	E_CELL_MANAGER_STATE.WAIT_GRIPPER1_CONTENT:
		IF rtOperatorChoice.Q AND xOperatorChoiceAllowed THEN
			IF uiOperatorChoice = UINT#1 THEN
				IF Config.uiTypeCount = UINT#1 THEN
					uiBlankPayloadType := UINT#1;
					IF xPrestartGripper2Occupied THEN
						eState := E_CELL_MANAGER_STATE.WAIT_GRIPPER2_CONTENT;
					ELSE
						xSafetyHomeRequired := FALSE;
						xStoppedPoseValid := FALSE;
						xRunning := TRUE;
						eState := E_CELL_MANAGER_STATE.PLAN_TARGET;
					END_IF;
				ELSE
					eState := E_CELL_MANAGER_STATE.WAIT_GRIPPER1_TYPE;
				END_IF;
			ELSIF uiOperatorChoice = UINT#2 THEN
				Diag.stWarning.uiCode := WRN_GRIPPER1_CONTENT;
				Diag.stWarning.udiSequence := Diag.stWarning.udiSequence + UDINT#1;
				IF Diag.stWarning.udiSequence = UDINT#0 THEN Diag.stWarning.udiSequence := UDINT#1; END_IF;
				eState := E_CELL_MANAGER_STATE.IDLE;
			ELSE
				Diag.stWarning.uiCode := WRN_OPERATOR_REPLY_REJECTED;
				Diag.stWarning.udiSequence := Diag.stWarning.udiSequence + UDINT#1;
				IF Diag.stWarning.udiSequence = UDINT#0 THEN Diag.stWarning.udiSequence := UDINT#1; END_IF;
				eState := E_CELL_MANAGER_STATE.IDLE;
			END_IF;
		END_IF;

	E_CELL_MANAGER_STATE.WAIT_GRIPPER1_TYPE:
		IF rtOperatorChoice.Q AND xOperatorChoiceAllowed THEN
			IF (uiOperatorChoice >= UINT#1)
			AND (uiOperatorChoice <= Config.uiTypeCount) THEN
				uiBlankPayloadType := uiOperatorChoice;
				IF xPrestartGripper2Occupied THEN
					eState := E_CELL_MANAGER_STATE.WAIT_GRIPPER2_CONTENT;
				ELSE
					xSafetyHomeRequired := FALSE;
					xStoppedPoseValid := FALSE;
					xRunning := TRUE;
					eState := E_CELL_MANAGER_STATE.PLAN_TARGET;
				END_IF;
			ELSE
				Diag.stWarning.uiCode := WRN_PAYLOAD_TYPE_CHOICE;
				Diag.stWarning.udiSequence := Diag.stWarning.udiSequence + UDINT#1;
				IF Diag.stWarning.udiSequence = UDINT#0 THEN Diag.stWarning.udiSequence := UDINT#1; END_IF;
				eState := E_CELL_MANAGER_STATE.IDLE;
			END_IF;
		END_IF;

	E_CELL_MANAGER_STATE.WAIT_GRIPPER2_CONTENT:
		IF rtOperatorChoice.Q AND xOperatorChoiceAllowed THEN
			IF uiOperatorChoice = UINT#2 THEN
				IF Config.uiTypeCount = UINT#1 THEN
					uiDetailPayloadType := UINT#1;
				ELSE
					eState := E_CELL_MANAGER_STATE.WAIT_GRIPPER2_TYPE;
				END_IF;
				IF (Config.uiTypeCount = UINT#1) AND xPrestartGripper1Occupied THEN
					IF uiOperatorMachineMask <> UINT#0 THEN
						eState := E_CELL_MANAGER_STATE.WAIT_START_MACHINE;
					ELSE
						// Нет пустого совместимого станка: это не тупик. После
						// идентификации обоих грузов планировщик сначала уложит деталь.
						xSafetyHomeRequired := FALSE;
						xStoppedPoseValid := FALSE;
						xRunning := TRUE;
						eState := E_CELL_MANAGER_STATE.PLAN_TARGET;
					END_IF;
				ELSIF Config.uiTypeCount = UINT#1 THEN
					xSafetyHomeRequired := FALSE;
					xStoppedPoseValid := FALSE;
					xRunning := TRUE;
					eState := E_CELL_MANAGER_STATE.PLAN_TARGET;
				END_IF;
			ELSIF uiOperatorChoice = UINT#1 THEN
				Diag.stWarning.uiCode := WRN_GRIPPER2_CONTENT;
				Diag.stWarning.udiSequence := Diag.stWarning.udiSequence + UDINT#1;
				IF Diag.stWarning.udiSequence = UDINT#0 THEN Diag.stWarning.udiSequence := UDINT#1; END_IF;
				eState := E_CELL_MANAGER_STATE.IDLE;
			ELSE
				Diag.stWarning.uiCode := WRN_OPERATOR_REPLY_REJECTED;
				Diag.stWarning.udiSequence := Diag.stWarning.udiSequence + UDINT#1;
				IF Diag.stWarning.udiSequence = UDINT#0 THEN Diag.stWarning.udiSequence := UDINT#1; END_IF;
				eState := E_CELL_MANAGER_STATE.IDLE;
			END_IF;
		END_IF;

	E_CELL_MANAGER_STATE.WAIT_GRIPPER2_TYPE:
		IF rtOperatorChoice.Q AND xOperatorChoiceAllowed THEN
			IF (uiOperatorChoice >= UINT#1)
			AND (uiOperatorChoice <= Config.uiTypeCount) THEN
				uiDetailPayloadType := uiOperatorChoice;
				IF xPrestartGripper1Occupied THEN
					IF uiOperatorMachineMask <> UINT#0 THEN
						eState := E_CELL_MANAGER_STATE.WAIT_START_MACHINE;
					ELSE
						xSafetyHomeRequired := FALSE;
						xStoppedPoseValid := FALSE;
						xRunning := TRUE;
						eState := E_CELL_MANAGER_STATE.PLAN_TARGET;
					END_IF;
				ELSE
					xSafetyHomeRequired := FALSE;
					xStoppedPoseValid := FALSE;
					xRunning := TRUE;
					eState := E_CELL_MANAGER_STATE.PLAN_TARGET;
				END_IF;
			ELSE
				Diag.stWarning.uiCode := WRN_PAYLOAD_TYPE_CHOICE;
				Diag.stWarning.udiSequence := Diag.stWarning.udiSequence + UDINT#1;
				IF Diag.stWarning.udiSequence = UDINT#0 THEN Diag.stWarning.udiSequence := UDINT#1; END_IF;
				eState := E_CELL_MANAGER_STATE.IDLE;
			END_IF;
		END_IF;

	E_CELL_MANAGER_STATE.WAIT_START_MACHINE:
		IF (uiDetailPayloadType < UINT#1)
		OR (uiDetailPayloadType > Config.uiTypeCount) THEN
			Diag.stWarning.uiCode := WRN_PAYLOAD_TYPE_CHOICE;
			Diag.stWarning.udiSequence := Diag.stWarning.udiSequence + UDINT#1;
			IF Diag.stWarning.udiSequence = UDINT#0 THEN Diag.stWarning.udiSequence := UDINT#1; END_IF;
			eState := E_CELL_MANAGER_STATE.IDLE;
		ELSIF stMagazineStatus.stTypeStatus.aiFreeSlot[uiDetailPayloadType] = SINT#0 THEN
			Diag.stWarning.uiCode := WRN_DETAIL_SLOT_REQUIRED;
			Diag.stWarning.udiSequence := Diag.stWarning.udiSequence + UDINT#1;
			IF Diag.stWarning.udiSequence = UDINT#0 THEN Diag.stWarning.udiSequence := UDINT#1; END_IF;
			eState := E_CELL_MANAGER_STATE.IDLE;
		ELSIF uiOperatorMachineMask = UINT#0 THEN
			// Пока оператор отвечал, пустой станок мог стать недоступен. Сохраняем
			// оба груза и передаём решение общему планировщику вместо отмены старта.
			xSafetyHomeRequired := FALSE;
			xStoppedPoseValid := FALSE;
			xRunning := TRUE;
			eState := E_CELL_MANAGER_STATE.PLAN_TARGET;
		ELSIF rtOperatorChoice.Q AND xOperatorChoiceAllowed THEN
			IF ((uiOperatorChoice = UINT#1) AND ((uiOperatorMachineMask AND UINT#1) <> UINT#0))
			OR ((uiOperatorChoice = UINT#2) AND ((uiOperatorMachineMask AND UINT#2) <> UINT#0))
			OR ((uiOperatorChoice = UINT#3) AND ((uiOperatorMachineMask AND UINT#4) <> UINT#0)) THEN
				uiSelectedMachine := uiOperatorChoice;
				uiSelectedType := uiBlankPayloadType;
				eMachineOperation := E_MACHINE_OPERATION.LOAD;
				xSafetyHomeRequired := FALSE;
				xStoppedPoseValid := FALSE;
				xRunning := TRUE;
				eState := E_CELL_MANAGER_STATE.ROUTE_TO_TARGET;
			ELSE
				Diag.stWarning.uiCode := WRN_START_MACHINE_CHOICE;
				Diag.stWarning.udiSequence := Diag.stWarning.udiSequence + UDINT#1;
				IF Diag.stWarning.udiSequence = UDINT#0 THEN Diag.stWarning.udiSequence := UDINT#1; END_IF;
				eState := E_CELL_MANAGER_STATE.IDLE;
			END_IF;
		END_IF;

	E_CELL_MANAGER_STATE.PLAN_TARGET:
		IF xStopRequested
		AND NOT stRobotStatus.xBusy
		AND NOT stMagazineStatus.xBusy THEN
			xRunning := FALSE;
			eState := E_CELL_MANAGER_STATE.IDLE;

		ELSIF PlanGeometry() THEN
			// Метод зафиксировал резерв или безопасное ожидание свободного ГК.
		ELSIF stRobotStatus.xBlankAvailable
		AND stRobotStatus.xDetailAvailable THEN
			// Два груза после аварийного восстановления — штатная ситуация. Сначала
			// ищем пустой готовый станок строго по типу заготовки. Если загрузить её
			// прямо сейчас некуда, освобождаем захват 2 операцией PUT.
			IF (uiBlankPayloadType < UINT#1)
			OR (uiBlankPayloadType > Config.uiTypeCount) THEN
				Error.dwErrorActive := Error.dwErrorActive OR ERR_MAGAZINE;
				eState := E_CELL_MANAGER_STATE.ERROR;
			ELSIF (uiDetailPayloadType < UINT#1)
			OR (uiDetailPayloadType > Config.uiTypeCount) THEN
				Error.dwErrorActive := Error.dwErrorActive OR ERR_MACHINE;
				eState := E_CELL_MANAGER_STATE.ERROR;
			ELSE
				uiCandidateMachine := UINT#0;
				FOR uiMachine := FIRST_MACHINE TO LAST_MACHINE DO
					IF (uiCandidateMachine = UINT#0)
					AND IsMachineCompatible(
						uiMachine := uiMachine,
						uiProductType := uiBlankPayloadType
					)
					AND astMachineStatus[uiMachine].xCanAcceptService
					AND (astMachineStatus[uiMachine].ePartState = E_PART_STATE.EMPTY) THEN
						uiCandidateMachine := uiMachine;
					END_IF;
				END_FOR;

				IF uiCandidateMachine > UINT#0 THEN
					uiSelectedMachine := uiCandidateMachine;
					uiSelectedType := uiBlankPayloadType;
					eMachineOperation := E_MACHINE_OPERATION.LOAD;
					xMachineServiceStarted := FALSE;
					eState := E_CELL_MANAGER_STATE.ROUTE_TO_TARGET;
				ELSIF (stMagazineStatus.stTypeStatus.aiFreeSlot[uiDetailPayloadType] > SINT#0)
				AND xMagazineReady THEN
					uiSelectedMachine := UINT#0;
					uiSelectedType := UINT#0;
					eMachineOperation := E_MACHINE_OPERATION.NONE;
					iTakeSlot := SINT#0;
					iTakeOriginSlot := SINT#0;
					iPutSlot := stMagazineStatus.stTypeStatus.aiFreeSlot[uiDetailPayloadType];
					eMagazineOperation := E_MAGAZINE_OPERATION.PUT;
					eState := E_CELL_MANAGER_STATE.MAGAZINE_EXECUTE;
				ELSE
					eState := E_CELL_MANAGER_STATE.WAIT_MAGAZINE;
				END_IF;
			END_IF;

		ELSIF stRobotStatus.xBlankAvailable THEN
			IF (uiBlankPayloadType < UINT#1)
			OR (uiBlankPayloadType > Config.uiTypeCount) THEN
				Error.dwErrorActive := Error.dwErrorActive OR ERR_MAGAZINE;
				eState := E_CELL_MANAGER_STATE.ERROR;
			ELSE
				uiSelectedType := uiBlankPayloadType;
				uiCandidateMachine := SelectMachineForHeldBlank(
					uiProductType := uiBlankPayloadType,
					uiCurrentMachine := uiSelectedMachine
				);
				IF uiCandidateMachine > UINT#0 THEN
					uiSelectedMachine := uiCandidateMachine;
					eState := E_CELL_MANAGER_STATE.ROUTE_TO_TARGET;
				ELSE
					uiSelectedMachine := UINT#0;
					eState := E_CELL_MANAGER_STATE.SELECT_FALLBACK;
				END_IF;
			END_IF;

		ELSIF stRobotStatus.xDetailAvailable THEN
			uiBlankPayloadType := UINT#0;
			IF (uiDetailPayloadType < UINT#1)
			OR (uiDetailPayloadType > Config.uiTypeCount) THEN
				Error.dwErrorActive := Error.dwErrorActive OR ERR_MACHINE;
				eState := E_CELL_MANAGER_STATE.ERROR;
			ELSIF NOT xMagazineReady THEN
				eState := E_CELL_MANAGER_STATE.WAIT_MAGAZINE;
			ELSE
				// При полной палете CHANGE сначала освобождает слот взятием заготовки.
				// Станок назначения может быть пустым, готовым к обмену или обрабатывать.
				iPutSlot := stMagazineStatus.stTypeStatus.aiFreeSlot[uiDetailPayloadType];
				uiCandidateMachine := SelectMachineBeforeTake();
				uiSelectedMachine := UINT#0;
				uiSelectedType := UINT#0;
				iTakeSlot := SINT#0;
				iTakeOriginSlot := SINT#0;
				eMachineOperation := E_MACHINE_OPERATION.NONE;

				// Закрытый или переходный первый захват исключает CHANGE, даже если
				// логический флаг груза сейчас снят.
				IF stRobotStatus.xGripper1Open
				AND (uiCandidateMachine >= FIRST_MACHINE)
				AND (uiCandidateMachine <= LAST_MACHINE) THEN
					uiSelectedMachine := uiCandidateMachine;
					uiSelectedType := Config.auiMachineType[uiSelectedMachine];
					IF (uiSelectedType >= UINT#1)
					AND (uiSelectedType <= Config.uiTypeCount) THEN
						iTakeSlot := stMagazineStatus.stTypeStatus.aiBlankSlot[uiSelectedType];
					END_IF;
				END_IF;

				// Индексы проверяются до обращения к карте секций. Обычный AND в
				// CODESYS не используется как защита динамического индекса массива.
				IF iPutSlot = SINT#0 THEN
					iPutSlot := iTakeSlot;
				END_IF;
				IF (iPutSlot >= SINT#1)
				AND (SINT_TO_UINT(iPutSlot) <= SINT_TO_UINT(GVL_CELL_SETTINGS.NumberDetail))
				AND (iTakeSlot >= SINT#1)
				AND (SINT_TO_UINT(iTakeSlot) <= SINT_TO_UINT(GVL_CELL_SETTINGS.NumberDetail)) THEN
					xChangePrepared := TRUE;
				END_IF;

				IF xChangePrepared THEN
					iTakeOriginSlot := iTakeSlot;
					eMagazineOperation := E_MAGAZINE_OPERATION.CHANGE;
					eState := E_CELL_MANAGER_STATE.MAGAZINE_EXECUTE;
				ELSE
					// Если следующую заготовку нельзя безопасно назначить, сначала
					// освобождаем второй захват и пересчитываем маршрут после PUT.
					uiSelectedMachine := UINT#0;
					uiSelectedType := UINT#0;
					iTakeSlot := SINT#0;
					iTakeOriginSlot := SINT#0;
					IF stMagazineStatus.stTypeStatus.aiFreeSlot[uiDetailPayloadType] > SINT#0 THEN
						iPutSlot := stMagazineStatus.stTypeStatus.aiFreeSlot[uiDetailPayloadType];
						eMagazineOperation := E_MAGAZINE_OPERATION.PUT;
						eState := E_CELL_MANAGER_STATE.MAGAZINE_EXECUTE;
					ELSE
						iPutSlot := SINT#0;
						eMagazineOperation := E_MAGAZINE_OPERATION.NONE;
						eState := E_CELL_MANAGER_STATE.WAIT_MAGAZINE;
					END_IF;
				END_IF;
			END_IF;

		ELSE
			uiBlankPayloadType := UINT#0;
			uiDetailPayloadType := UINT#0;
			uiCandidateMachine := SelectMachineBeforeTake();
			IF uiCandidateMachine > UINT#0 THEN
				IF NOT xMagazineReady THEN
					eState := E_CELL_MANAGER_STATE.WAIT_MAGAZINE;
				ELSE
					uiSelectedMachine := uiCandidateMachine;
					uiSelectedType := Config.auiMachineType[uiSelectedMachine];
					iTakeSlot := stMagazineStatus.stTypeStatus.aiBlankSlot[uiSelectedType];
					iTakeOriginSlot := iTakeSlot;
					iPutSlot := SINT#0;
					eMachineOperation := E_MACHINE_OPERATION.NONE;
					eMagazineOperation := E_MAGAZINE_OPERATION.TAKE;
					eState := E_CELL_MANAGER_STATE.MAGAZINE_EXECUTE;
				END_IF;
			ELSE
				// Заготовок в магазине нет — выбираем готовую деталь для отдельной выгрузки.
				uiCandidateMachine := SelectMachineForUnload(uiCurrentMachine := UINT#0);
				IF uiCandidateMachine > UINT#0 THEN
					uiSelectedMachine := uiCandidateMachine;
					uiSelectedType := Config.auiMachineType[uiSelectedMachine];
					eMachineOperation := E_MACHINE_OPERATION.UNLOAD;
					xMachineServiceStarted := FALSE;
					iTakeSlot := SINT#0;
					iPutSlot := SINT#0;
					IF xMagazineReady THEN
						eState := E_CELL_MANAGER_STATE.ROUTE_TO_TARGET;
					ELSE
						eState := E_CELL_MANAGER_STATE.WAIT_MAGAZINE;
					END_IF;
				ELSE
					IF stMagazineStatus.xFinished THEN
						eState := E_CELL_MANAGER_STATE.WAIT_MAGAZINE;
					ELSE
						eState := E_CELL_MANAGER_STATE.WAIT_TARGET;
					END_IF;
				END_IF;
			END_IF;
		END_IF;

	E_CELL_MANAGER_STATE.MAGAZINE_EXECUTE:
		IF xGeometryHeld AND (uiGeometryMachine >= UINT#1) AND (uiGeometryMachine <= UINT#3)
		AND (stMagazineStatus.udiProducedPartsTotal <> udiGeometryMagazineCounter)
		AND NOT stRobotStatus.xDetailAvailable AND stRobotStatus.xGripper2Open THEN
			GVL_GEOMETRY_CONTROL.astCalls[uiGeometryMachine].uiState := UINT#5;
			GVL_GEOMETRY_CONTROL.astCalls[uiGeometryMachine].uiReason := uiGeometryBypassReason;
			GVL_GEOMETRY_CONTROL.astCalls[uiGeometryMachine].uiMagazine := uiActiveMagazine;
			GVL_GEOMETRY_CONTROL.astCalls[uiGeometryMachine].uiSlot := SINT_TO_UINT(iPutSlot);
			IF GVL_TWO_PALLET.uiMode = UINT#1 THEN
				GVL_GEOMETRY_CONTROL.astCalls[uiGeometryMachine].uiPallet := GVL_TWO_PALLET.astStatus[uiActiveMagazine].uiRobotPallet;
			END_IF;
			F_GEOMETRY_EVENT(Call := GVL_GEOMETRY_CONTROL.astCalls[uiGeometryMachine]);
			GVL_GEOMETRY_CONTROL.stCellWarning.uiCode := UINT#50;
			GVL_GEOMETRY_CONTROL.stCellWarning.udiSequence := GVL_GEOMETRY_CONTROL.stCellWarning.udiSequence + UDINT#1;
			xGeometryHeld := FALSE; uiGeometryMachine := UINT#0;
		END_IF;
		Command.stMagazine.xExecute := TRUE;
		IF (eMagazineOperation = E_MAGAZINE_OPERATION.NONE) THEN
			Error.dwErrorActive := Error.dwErrorActive OR ERR_MAGAZINE;
			eState := E_CELL_MANAGER_STATE.ERROR;
		END_IF;

		IF stMagazineStatus.xError THEN
			Command.stMagazine.xExecute := FALSE;
			IF stMagazineStatus.xRobotStopRequired THEN
				xSafetyHomeRequired := TRUE;
				xStoppedPoseValid := FALSE;
				Error.dwErrorActive := Error.dwErrorActive OR ERR_MAGAZINE;
				eState := E_CELL_MANAGER_STATE.ERROR;
			ELSE
				xRunning := FALSE;
				eState := E_CELL_MANAGER_STATE.IDLE;
			END_IF;
		ELSIF stRobotStatus.xError THEN
			Error.dwErrorActive := Error.dwErrorActive OR ERR_ROBOT;
			eState := E_CELL_MANAGER_STATE.ERROR;
		ELSIF stMagazineStatus.xDone THEN
			eState := E_CELL_MANAGER_STATE.RELEASE_MAGAZINE;
		END_IF;

	E_CELL_MANAGER_STATE.RELEASE_MAGAZINE:
		IF stMagazineStatus.xError THEN
			IF stMagazineStatus.xRobotStopRequired THEN
				xSafetyHomeRequired := TRUE;
				xStoppedPoseValid := FALSE;
				Error.dwErrorActive := Error.dwErrorActive OR ERR_MAGAZINE;
				eState := E_CELL_MANAGER_STATE.ERROR;
			ELSE
				xRunning := FALSE;
				eState := E_CELL_MANAGER_STATE.IDLE;
			END_IF;
		ELSIF NOT stMagazineStatus.xBusy
		AND NOT stMagazineStatus.xDone THEN
			CASE eMagazineOperation OF
				E_MAGAZINE_OPERATION.TAKE:
					uiBlankPayloadType := uiSelectedType;
				E_MAGAZINE_OPERATION.PUT:
					uiDetailPayloadType := UINT#0;
				E_MAGAZINE_OPERATION.CHANGE:
					uiDetailPayloadType := UINT#0;
					uiBlankPayloadType := uiSelectedType;
				E_MAGAZINE_OPERATION.RETURN_BLANK:
					uiBlankPayloadType := UINT#0;
					uiSelectedType := UINT#0;
					iTakeOriginSlot := SINT#0;
					iTakeSlot := SINT#0;
					iPutSlot := SINT#0;
			END_CASE;
			eMagazineOperation := E_MAGAZINE_OPERATION.NONE;
			eState := E_CELL_MANAGER_STATE.PLAN_TARGET;
		END_IF;

	E_CELL_MANAGER_STATE.ROUTE_TO_TARGET:
		IF eMachineOperation = E_MACHINE_OPERATION.UNLOAD THEN
			IF stRobotStatus.eCurrentPoint = astMachineStatus[uiSelectedMachine].eAbovePoint THEN
				eState := E_CELL_MANAGER_STATE.WAIT_TARGET;
			ELSE
				Command.stRobot.xExecute := TRUE;
				Command.stRobot.eAction := E_ROBOT_ACTION.MOVE_TO_POINT;
				Command.stRobot.eSetPoint := astMachineStatus[uiSelectedMachine].eAbovePoint;
				IF stRobotStatus.xDone THEN
					xReselectAfterRobotRelease := FALSE;
					eState := E_CELL_MANAGER_STATE.RELEASE_ROBOT_COMMAND;
				END_IF;
			END_IF;
		ELSE
			IF (uiSelectedMachine >= FIRST_MACHINE)
			AND (uiSelectedMachine <= LAST_MACHINE) THEN
				RaisePayloadRouteWarning(
					uiPayloadType := uiBlankPayloadType,
					uiDestinationType := Config.auiMachineType[uiSelectedMachine]
				);
			END_IF;
			IF NOT IsMachineCompatible(
				uiMachine := uiSelectedMachine,
				uiProductType := uiBlankPayloadType
			) THEN
				xReselectAfterRobotRelease := TRUE;
				eState := E_CELL_MANAGER_STATE.RELEASE_ROBOT_COMMAND;
			ELSIF stRobotStatus.eCurrentPoint = astMachineStatus[uiSelectedMachine].eAbovePoint THEN
				eState := E_CELL_MANAGER_STATE.WAIT_TARGET;
			ELSE
				Command.stRobot.xExecute := TRUE;
				Command.stRobot.eAction := E_ROBOT_ACTION.MOVE_TO_POINT;
				Command.stRobot.eSetPoint := astMachineStatus[uiSelectedMachine].eAbovePoint;
				IF stRobotStatus.xDone THEN
					xReselectAfterRobotRelease := FALSE;
					eState := E_CELL_MANAGER_STATE.RELEASE_ROBOT_COMMAND;
				END_IF;
			END_IF;
		END_IF;

	E_CELL_MANAGER_STATE.RELEASE_ROBOT_COMMAND:
		IF stRobotStatus.xError THEN
			Error.dwErrorActive := Error.dwErrorActive OR ERR_ROBOT;
			eState := E_CELL_MANAGER_STATE.ERROR;
		ELSIF NOT stRobotStatus.xBusy
		AND NOT stRobotStatus.xDone THEN
			IF eMachineOperation = E_MACHINE_OPERATION.UNLOAD THEN
				eState := E_CELL_MANAGER_STATE.WAIT_TARGET;
			ELSIF xReselectAfterRobotRelease THEN
				xReselectAfterRobotRelease := FALSE;
				eState := E_CELL_MANAGER_STATE.SELECT_FALLBACK;
			ELSIF IsMachineCompatible(
				uiMachine := uiSelectedMachine,
				uiProductType := uiBlankPayloadType
			) THEN
				eState := E_CELL_MANAGER_STATE.WAIT_TARGET;
			ELSE
				eState := E_CELL_MANAGER_STATE.SELECT_FALLBACK;
			END_IF;
		END_IF;

	E_CELL_MANAGER_STATE.WAIT_TARGET:
		IF xStopRequested
		AND NOT stRobotStatus.xBusy THEN
			xRunning := FALSE;
			eState := E_CELL_MANAGER_STATE.IDLE;
		ELSIF (eMachineOperation = E_MACHINE_OPERATION.UNLOAD)
		AND NOT stRobotStatus.xBlankAvailable
		AND NOT stRobotStatus.xDetailAvailable THEN
			uiCandidateMachine := SelectMachineForUnload(uiCurrentMachine := uiSelectedMachine);
			IF uiCandidateMachine = UINT#0 THEN
				uiSelectedMachine := UINT#0;
				uiSelectedType := UINT#0;
				eMachineOperation := E_MACHINE_OPERATION.NONE;
				IF stMagazineStatus.xFinished THEN
					eState := E_CELL_MANAGER_STATE.WAIT_MAGAZINE;
				ELSE
					eState := E_CELL_MANAGER_STATE.PLAN_TARGET;
				END_IF;
			ELSIF uiCandidateMachine <> uiSelectedMachine THEN
				uiSelectedMachine := uiCandidateMachine;
				uiSelectedType := Config.auiMachineType[uiSelectedMachine];
				eState := E_CELL_MANAGER_STATE.ROUTE_TO_TARGET;
			ELSIF stRobotStatus.eCurrentPoint <> astMachineStatus[uiSelectedMachine].eAbovePoint THEN
				eState := E_CELL_MANAGER_STATE.ROUTE_TO_TARGET;
			ELSIF astMachineStatus[uiSelectedMachine].xCanAcceptService
			AND astMachineStatus[uiSelectedMachine].xServiceRequired
			AND (astMachineStatus[uiSelectedMachine].ePartState = E_PART_STATE.LOADED)
			AND (astMachineStatus[uiSelectedMachine].ePartType = E_PART_TYPE.DETAIL) THEN
				xMachineServiceStarted := FALSE;
				eState := E_CELL_MANAGER_STATE.SERVICE_TARGET;
			END_IF;
		ELSIF stRobotStatus.xBlankAvailable
		AND stRobotStatus.xDetailAvailable THEN
			// Выбранная пустая цель могла стать недоступной по дороге. Обслуживаем
			// только всё ещё пустой совместимый станок; иначе перепланируем через PUT.
			IF (uiSelectedMachine >= FIRST_MACHINE)
			AND (uiSelectedMachine <= LAST_MACHINE) THEN
				IF IsMachineCompatible(
					uiMachine := uiSelectedMachine,
					uiProductType := uiBlankPayloadType
				)
				AND (stRobotStatus.eCurrentPoint = astMachineStatus[uiSelectedMachine].eAbovePoint)
				AND astMachineStatus[uiSelectedMachine].xCanAcceptService
				AND (astMachineStatus[uiSelectedMachine].ePartState = E_PART_STATE.EMPTY) THEN
					eMachineOperation := E_MACHINE_OPERATION.LOAD;
					xMachineServiceStarted := FALSE;
					eState := E_CELL_MANAGER_STATE.SERVICE_TARGET;
				ELSE
					eState := E_CELL_MANAGER_STATE.PLAN_TARGET;
				END_IF;
			ELSE
				eState := E_CELL_MANAGER_STATE.PLAN_TARGET;
			END_IF;
		ELSIF stRobotStatus.xBlankAvailable THEN
			uiCandidateMachine := SelectMachineForHeldBlank(
				uiProductType := uiBlankPayloadType,
				uiCurrentMachine := uiSelectedMachine
			);
			IF uiCandidateMachine = UINT#0 THEN
				eState := E_CELL_MANAGER_STATE.SELECT_FALLBACK;
			ELSIF uiCandidateMachine <> uiSelectedMachine THEN
				uiSelectedMachine := uiCandidateMachine;
				eState := E_CELL_MANAGER_STATE.ROUTE_TO_TARGET;
			ELSIF stRobotStatus.eCurrentPoint <> astMachineStatus[uiSelectedMachine].eAbovePoint THEN
				eState := E_CELL_MANAGER_STATE.ROUTE_TO_TARGET;
			ELSIF astMachineStatus[uiSelectedMachine].xCanAcceptService
			AND astMachineStatus[uiSelectedMachine].xServiceRequired THEN
				eMachineOperation := astMachineStatus[uiSelectedMachine].eRecommendedOperation;
				axMachineStartPending[uiSelectedMachine] := FALSE;
				xMachineServiceStarted := FALSE;
				eState := E_CELL_MANAGER_STATE.SERVICE_TARGET;
			END_IF;
		ELSIF stRobotStatus.xDetailAvailable THEN
			// Готовая деталь в захвате обслуживается через общий план PUT.
			eState := E_CELL_MANAGER_STATE.PLAN_TARGET;
		ELSE
			uiCandidateMachine := SelectMachineBeforeTake();
			IF uiCandidateMachine > UINT#0 THEN
				eState := E_CELL_MANAGER_STATE.PLAN_TARGET;
			ELSE
				// В магазине нет заготовки: ожидаем готовую деталь станка,
				// которую можно выгрузить в свободный слот.
				uiCandidateMachine := SelectMachineForUnload(uiCurrentMachine := uiSelectedMachine);
				IF uiCandidateMachine > UINT#0 THEN
					uiSelectedMachine := uiCandidateMachine;
					uiSelectedType := Config.auiMachineType[uiSelectedMachine];
					eMachineOperation := E_MACHINE_OPERATION.UNLOAD;
					xMachineServiceStarted := FALSE;
					iTakeSlot := SINT#0;
					iPutSlot := SINT#0;
					IF xMagazineReady THEN
						eState := E_CELL_MANAGER_STATE.ROUTE_TO_TARGET;
					ELSE
						eState := E_CELL_MANAGER_STATE.WAIT_MAGAZINE;
					END_IF;
				ELSIF stMagazineStatus.xFinished THEN
					eState := E_CELL_MANAGER_STATE.WAIT_MAGAZINE;
				END_IF;
			END_IF;
		END_IF;

	E_CELL_MANAGER_STATE.SERVICE_TARGET:
		IF (uiSelectedMachine < FIRST_MACHINE)
		OR (uiSelectedMachine > LAST_MACHINE) THEN
			Error.dwErrorActive := Error.dwErrorActive OR ERR_MACHINE;
			eState := E_CELL_MANAGER_STATE.ERROR;
		ELSIF NOT xMachineServiceStarted AND NOT astMachineStatus[uiSelectedMachine].xBusy
		AND (eMachineOperation <> E_MACHINE_OPERATION.LOAD)
		AND axGeometryUnloadBlocked[uiSelectedMachine] THEN
			// До запуска рецепта повторно проверяем свободный ГК и очередь вызовов.
			// Деталь остаётся в патроне; ищем другую работу без команды станку.
			eState := E_CELL_MANAGER_STATE.SELECT_FALLBACK;
		ELSIF NOT xMachineServiceStarted
		AND (eMachineOperation <> E_MACHINE_OPERATION.UNLOAD)
		AND NOT IsMachineCompatible(
			uiMachine := uiSelectedMachine,
			uiProductType := uiBlankPayloadType
		) THEN
			RaisePayloadRouteWarning(
				uiPayloadType := uiBlankPayloadType,
				uiDestinationType := Config.auiMachineType[uiSelectedMachine]
			);
			eState := E_CELL_MANAGER_STATE.SELECT_FALLBACK;
		ELSE
			IF NOT xMachineServiceStarted AND NOT stRobotStatus.xDetailAvailable THEN xGeometryDetailCounted := FALSE; END_IF;
			IF stRobotStatus.xDetailAvailable AND NOT xGeometryDetailCounted
			AND ((eMachineOperation = E_MACHINE_OPERATION.CHANGE) OR (eMachineOperation = E_MACHINE_OPERATION.UNLOAD)) THEN
				xGeometryHeld := F_GEOMETRY_TAKE_DETAIL(uiMachine := uiSelectedMachine, uiProductType := Config.auiMachineType[uiSelectedMachine]);
				IF xGeometryHeld THEN uiGeometryMachine := uiSelectedMachine; uiGeometryBypassReason := UINT#0; END_IF;
				xGeometryDetailCounted := TRUE;
			END_IF;
			// Тип детали передаётся в FB_ROBOT сразу после фактического закрытия
			// второго захвата, а не после полного выхода робота из станка.
			IF stRobotStatus.xDetailAvailable
			AND ((eMachineOperation = E_MACHINE_OPERATION.CHANGE)
				OR (eMachineOperation = E_MACHINE_OPERATION.UNLOAD)) THEN
				uiDetailPayloadType := Config.auiMachineType[uiSelectedMachine];
			END_IF;
			IF eMachineOperation <> E_MACHINE_OPERATION.UNLOAD THEN
				RaisePayloadRouteWarning(
					uiPayloadType := uiBlankPayloadType,
					uiDestinationType := Config.auiMachineType[uiSelectedMachine]
				);
			END_IF;
			Command.axMachineExecute[uiSelectedMachine] := TRUE;
			IF astMachineStatus[uiSelectedMachine].xBusy THEN
				xMachineServiceStarted := TRUE;
			END_IF;

			IF astMachineStatus[uiSelectedMachine].xServiceRejected THEN
				Command.axMachineExecute[uiSelectedMachine] := FALSE;
				xMachineServiceStarted := FALSE;
				eState := E_CELL_MANAGER_STATE.SELECT_FALLBACK;
			ELSIF astMachineStatus[uiSelectedMachine].xError THEN
				Command.axMachineExecute[uiSelectedMachine] := FALSE;
				xMachineServiceStarted := FALSE;
				// ROBOT_STOP уже публикует сам станок и обрабатывает FB_ROBOT.
				// Локальная ошибка без робота просто исключает станок из маршрута.
				eState := E_CELL_MANAGER_STATE.SELECT_FALLBACK;
			ELSIF stRobotStatus.xError THEN
				Error.dwErrorActive := Error.dwErrorActive OR ERR_ROBOT;
				eState := E_CELL_MANAGER_STATE.ERROR;
			ELSIF astMachineStatus[uiSelectedMachine].xRobotReleased THEN
				// Вызов мог прийти после взятия детали, пока робот ещё менял заготовку.
				// Последняя проверка — после подтверждённого выхода, до сброса станка.
				// Только state 1: F_GEOMETRY_TAKE_DETAIL не считает выгрузку повторно
				// и привязывает ожидающий вызов лишь при его первом месте в FIFO.
				IF NOT xGeometryHeld AND stRobotStatus.xDetailAvailable
				AND ((eMachineOperation = E_MACHINE_OPERATION.CHANGE)
					OR (eMachineOperation = E_MACHINE_OPERATION.UNLOAD))
				AND (GVL_GEOMETRY_CONTROL.astCalls[uiSelectedMachine].uiState = UINT#1) THEN
					xGeometryHeld := F_GEOMETRY_TAKE_DETAIL(uiMachine := uiSelectedMachine, uiProductType := Config.auiMachineType[uiSelectedMachine]);
					IF xGeometryHeld THEN uiGeometryMachine := uiSelectedMachine; uiGeometryBypassReason := UINT#0; END_IF;
				END_IF;
				IF (eMachineOperation = E_MACHINE_OPERATION.LOAD)
				OR (eMachineOperation = E_MACHINE_OPERATION.CHANGE) THEN
					axMachineStartPending[uiSelectedMachine] := TRUE;
				END_IF;
				uiBlankPayloadType := UINT#0;
				IF (eMachineOperation = E_MACHINE_OPERATION.CHANGE)
				OR (eMachineOperation = E_MACHINE_OPERATION.UNLOAD) THEN
					uiDetailPayloadType := Config.auiMachineType[uiSelectedMachine];
				END_IF;
				uiSelectedMachine := UINT#0;
				uiSelectedType := UINT#0;
				xMachineServiceStarted := FALSE;
				eMachineOperation := E_MACHINE_OPERATION.NONE;
				eState := E_CELL_MANAGER_STATE.PLAN_TARGET;
			END_IF;
		END_IF;

	E_CELL_MANAGER_STATE.MACHINE_FAULT_STOP:
		// Удерживаем штатную остановку до полного освобождения Motion-слоя.
		// Первичная MachineAlarm/Timeout остаётся активной только в FB_MACHINE.
		Command.stRobot.xStop := stRobotStatus.xBusy OR xMotionBusy;
		IF NOT stRobotStatus.xBusy AND NOT xMotionBusy THEN
			xRunning := FALSE;
			xStopRequested := FALSE;
			xMachineServiceStarted := FALSE;
			xReselectAfterRobotRelease := FALSE;
			IF (uiSelectedMachine >= FIRST_MACHINE)
			AND (uiSelectedMachine <= LAST_MACHINE) THEN
				axMachineStartPending[uiSelectedMachine] := FALSE;
			END_IF;
			uiSelectedMachine := UINT#0;
			uiSelectedType := UINT#0;
			eMachineOperation := E_MACHINE_OPERATION.NONE;
			eState := E_CELL_MANAGER_STATE.IDLE;
		END_IF;

	E_CELL_MANAGER_STATE.SELECT_FALLBACK:
		IF xStopRequested
		AND NOT stRobotStatus.xBusy
		AND NOT stMagazineStatus.xBusy THEN
			xRunning := FALSE;
			eState := E_CELL_MANAGER_STATE.IDLE;
		ELSIF stRobotStatus.xDetailAvailable THEN
			// RETURN_BLANK запрещён при занятом захвате 2. Общий план сначала
			// попробует другой пустой станок, затем освободит готовую деталь через PUT.
			eState := E_CELL_MANAGER_STATE.PLAN_TARGET;
		ELSIF (uiBlankPayloadType < UINT#1)
		OR (uiBlankPayloadType > Config.uiTypeCount) THEN
			Error.dwErrorActive := Error.dwErrorActive OR ERR_MAGAZINE;
			eState := E_CELL_MANAGER_STATE.ERROR;
		ELSE
			uiCandidateMachine := SelectMachineForHeldBlank(
				uiProductType := uiBlankPayloadType,
				uiCurrentMachine := uiSelectedMachine
			);
		END_IF;
		IF (eState = E_CELL_MANAGER_STATE.SELECT_FALLBACK)
		AND (uiCandidateMachine > UINT#0) THEN
			uiSelectedMachine := uiCandidateMachine;
			uiSelectedType := uiBlankPayloadType;
			eState := E_CELL_MANAGER_STATE.ROUTE_TO_TARGET;
		ELSIF eState = E_CELL_MANAGER_STATE.SELECT_FALLBACK THEN
			uiSelectedMachine := UINT#0;
			eMachineOperation := E_MACHINE_OPERATION.NONE;
			eMagazineOperation := E_MAGAZINE_OPERATION.NONE;
			iPutSlot := SINT#0;
			IF NOT CanReturnHeldBlank() THEN
				// Один тип либо нет полезной работы другого типа: сохраняем
				// заготовку. WAIT_MAGAZINE заново проверяет маршруты без Start.
				eState := E_CELL_MANAGER_STATE.WAIT_MAGAZINE;
			ELSE
				// Исходный слот гарантированно освободился после подтверждённой TAKE.
				IF (iTakeOriginSlot >= SINT#1)
				AND (SINT_TO_UINT(iTakeOriginSlot) <= SINT_TO_UINT(GVL_CELL_SETTINGS.NumberDetail)) THEN
					iPutSlot := iTakeOriginSlot;
				END_IF;
				IF iPutSlot = SINT#0 THEN
					iPutSlot := stMagazineStatus.stTypeStatus.aiFreeSlot[uiBlankPayloadType];
				END_IF;
				IF (iPutSlot > SINT#0) AND xMagazineReady THEN
					eMagazineOperation := E_MAGAZINE_OPERATION.RETURN_BLANK;
					eState := E_CELL_MANAGER_STATE.MAGAZINE_EXECUTE;
				ELSE
					eState := E_CELL_MANAGER_STATE.WAIT_MAGAZINE;
				END_IF;
			END_IF;
		END_IF;

	E_CELL_MANAGER_STATE.WAIT_MAGAZINE:
		IF xStopRequested
		AND NOT stMagazineStatus.xBusy
		AND NOT stRobotStatus.xBusy THEN
			xRunning := FALSE;
			eState := E_CELL_MANAGER_STATE.IDLE;
		ELSIF stMagazineStatus.xError THEN
			IF stMagazineStatus.xRobotStopRequired THEN
				Error.dwErrorActive := Error.dwErrorActive OR ERR_MAGAZINE;
				eState := E_CELL_MANAGER_STATE.ERROR;
			ELSE
				xRunning := FALSE;
				eState := E_CELL_MANAGER_STATE.IDLE;
			END_IF;
		ELSIF stRobotStatus.xBlankAvailable
		AND stRobotStatus.xDetailAvailable THEN
			IF (uiBlankPayloadType < UINT#1)
			OR (uiBlankPayloadType > Config.uiTypeCount) THEN
				Error.dwErrorActive := Error.dwErrorActive OR ERR_MAGAZINE;
				eState := E_CELL_MANAGER_STATE.ERROR;
			ELSIF (uiDetailPayloadType < UINT#1)
			OR (uiDetailPayloadType > Config.uiTypeCount) THEN
				Error.dwErrorActive := Error.dwErrorActive OR ERR_MACHINE;
				eState := E_CELL_MANAGER_STATE.ERROR;
			ELSIF (uiOperatorMachineMask <> UINT#0)
			OR ((stMagazineStatus.stTypeStatus.aiFreeSlot[uiDetailPayloadType] > SINT#0)
				AND xMagazineReady) THEN
				eState := E_CELL_MANAGER_STATE.PLAN_TARGET;
			END_IF;
		ELSIF stRobotStatus.xBlankAvailable THEN
			IF (uiBlankPayloadType < UINT#1)
			OR (uiBlankPayloadType > Config.uiTypeCount) THEN
				Error.dwErrorActive := Error.dwErrorActive OR ERR_MAGAZINE;
				eState := E_CELL_MANAGER_STATE.ERROR;
			ELSE
				IF (SelectMachineForHeldBlank(
					uiProductType := uiBlankPayloadType,
					uiCurrentMachine := uiSelectedMachine
				) > UINT#0)
				OR CanReturnHeldBlank() THEN
					eState := E_CELL_MANAGER_STATE.SELECT_FALLBACK;
				END_IF;
			END_IF;
		ELSIF stRobotStatus.xDetailAvailable THEN
			IF (uiDetailPayloadType < UINT#1)
			OR (uiDetailPayloadType > Config.uiTypeCount) THEN
				Error.dwErrorActive := Error.dwErrorActive OR ERR_MACHINE;
				eState := E_CELL_MANAGER_STATE.ERROR;
			ELSE
				IF ((stMagazineStatus.stTypeStatus.aiFreeSlot[uiDetailPayloadType] > SINT#0)
					OR xActiveMagazineCanExchangeDetail)
				AND xMagazineReady THEN
					eState := E_CELL_MANAGER_STATE.PLAN_TARGET;
				END_IF;
			END_IF;
		ELSE
			uiCandidateMachine := SelectMachineBeforeTake();
			IF uiCandidateMachine = UINT#0 THEN
				uiCandidateMachine := SelectMachineForUnload(uiCurrentMachine := uiSelectedMachine);
			END_IF;
			IF uiCandidateMachine > UINT#0 THEN
				IF xMagazineReady THEN
					eState := E_CELL_MANAGER_STATE.PLAN_TARGET;
				ELSE
					eState := E_CELL_MANAGER_STATE.WAIT_MAGAZINE;
				END_IF;
			END_IF;
		END_IF;

	E_CELL_MANAGER_STATE.GEOMETRY_WAIT_FREE,
	E_CELL_MANAGER_STATE.GEOMETRY_DELIVER,
	E_CELL_MANAGER_STATE.GEOMETRY_RELEASE_COMMAND:
		RunGeometryRoute();

	E_CELL_MANAGER_STATE.ERROR:
		xRunning := FALSE;
		IF stRobotStatus.xBusy THEN
			Command.stRobot.xStop := TRUE;
		END_IF;
		IF stMagazineStatus.xBusy THEN
			Command.stMagazine.xStop := TRUE;
		END_IF;
		xResetAllowed := NOT xGlobalError
			AND NOT stRobotStatus.xBusy
			AND NOT stMagazineStatus.xBusy
			AND NOT xAnyMachineBusy
			AND NOT xMotionBusy;
		IF xReset AND xResetAllowed THEN
			Error.dwErrorLast := Error.dwErrorActive;
			Error.dwErrorActive := DWORD#0;
			IF NOT stRobotStatus.xBlankAvailable THEN
				uiBlankPayloadType := UINT#0;
			END_IF;
			IF NOT stRobotStatus.xDetailAvailable THEN
				uiDetailPayloadType := UINT#0;
			END_IF;
			eState := E_CELL_MANAGER_STATE.IDLE;
		END_IF;

	E_CELL_MANAGER_STATE.TEST_ABORT_STOP:
		xStopRequested := TRUE;
		Command.stRobot.xStop := TRUE;
		Command.stMagazine.xStop := TRUE;
		FOR uiMachine := FIRST_MACHINE TO LAST_MACHINE DO
			Command.axMachineExecute[uiMachine] := FALSE;
		END_FOR;
		IF NOT stRobotStatus.xBusy
		AND NOT xMotionBusy
		AND NOT stMagazineStatus.xBusy THEN
			xRunning := FALSE;
			xStopRequested := FALSE;
			xMachineServiceStarted := FALSE;
			xReselectAfterRobotRelease := FALSE;
			uiSelectedMachine := UINT#0;
			uiSelectedType := UINT#0;
			eMachineOperation := E_MACHINE_OPERATION.NONE;
			eMagazineOperation := E_MAGAZINE_OPERATION.NONE;
			eState := E_CELL_MANAGER_STATE.IDLE;
		END_IF;
END_CASE;

// Фиксируем позу только после завершённой штатной остановки или нормального
// окончания цикла. Аварийный переход оставляет xSafetyHomeRequired активным.
IF xWasRunning
AND NOT xRunning
AND (eState = E_CELL_MANAGER_STATE.IDLE)
AND NOT xSafetyHomeRequired THEN
	lrStoppedPoseX := lrRobotActualX;
	lrStoppedPoseY := lrRobotActualY;
	lrStoppedPoseZ := lrRobotActualZ;
	xStoppedPoseValid := TRUE;
END_IF;
xWasRunning := xRunning;

IF eState <> E_CELL_MANAGER_STATE.ERROR THEN
	xResetAllowed := FALSE;
END_IF;

Status.xMagazineExchangeAllowed := NOT xStopRequested
	AND ((eState = E_CELL_MANAGER_STATE.IDLE) OR (eState = E_CELL_MANAGER_STATE.PLAN_TARGET)
		OR (eState = E_CELL_MANAGER_STATE.WAIT_TARGET) OR (eState = E_CELL_MANAGER_STATE.WAIT_MAGAZINE));
Status.xRunning := xRunning;
Status.xStopPending := xStopRequested AND xRunning;
Status.xBusy := xRunning
	AND (eState <> E_CELL_MANAGER_STATE.IDLE)
	AND (eState <> E_CELL_MANAGER_STATE.ERROR);
Status.xWaitingMachine := (eState = E_CELL_MANAGER_STATE.WAIT_TARGET)
	OR (eState = E_CELL_MANAGER_STATE.SELECT_FALLBACK);
Status.xWaitingMagazine := eState = E_CELL_MANAGER_STATE.WAIT_MAGAZINE;
Status.xError := eState = E_CELL_MANAGER_STATE.ERROR;
Status.xReadyToStart := xReadyToStart;
Status.xStartAllowed := xReadyToStart
	OR (xRunning
		AND xStopRequested
		AND NOT xManual
		AND (eState <> E_CELL_MANAGER_STATE.MACHINE_FAULT_STOP));
Status.xStopAllowed := xRunning AND NOT xStopRequested;
Status.xResetAllowed := xResetAllowed;
// Ручной режим нельзя включить поверх работающего автоматического цикла.
// xManual уже отфильтрован до вызова FB, но это же условие публикуется HMI.
Status.xManualAllowed := NOT xRunning OR xGlobalError;
// В общей аварии оператору оставляем только ручное восстановление.
Status.xAutomaticAllowed := NOT xGlobalError AND NOT xIoEmergencyStopActive;
Status.xDrivesReady := xDrivesReady;
Status.xRobotReady := xRobotReady;
Status.xMagazineReady := xMagazineReady;
Status.xSafetyHomeRequired := xSafetyHomeRequired;
Status.xRobotAtSafetyHome := xRobotAtSafetyHome;
Status.xStartCheckCellIdle := xStartCheckCellIdle;
Status.xStartCheckAutomaticMode := xStartCheckAutomaticMode;
Status.xStartCheckNoBlockingError := xStartCheckNoBlockingError;
Status.xStartCheckRobotInterfaceReady := xStartCheckRobotInterfaceReady;
Status.xStartCheckConfigurationValid := xStartCheckConfigurationValid;
Status.xStartCheckPointsConfigured := xStartCheckPointsConfigured;
Status.xStartCheckDrivesReady := xStartCheckDrivesReady;
Status.xStartCheckRobotReady := xStartCheckRobotReady;
Status.xStartCheckMagazineReady := xStartCheckMagazineReady;
Status.xStartCheckTaskAvailable := xStartCheckTaskAvailable;
Status.xStartCheckSafetyHome := xStartCheckSafetyHome;
Status.xStartCheckSafety := xStartCheckSafety;
Status.uiStartConditionsMet := uiStartConditionsMet;
Status.uiStartConditionsTotal := UINT#12;
Status.uiReadyMachines := uiReadyMachines;
Status.uiSelectedMachine := uiSelectedMachine;
Status.uiActiveMagazine := uiActiveMagazine;
Status.eMagazineOperation := eMagazineOperation;
CASE eState OF
	E_CELL_MANAGER_STATE.WAIT_GRIPPER1_CONTENT: uiOperatorPrompt := UINT#1;
	E_CELL_MANAGER_STATE.WAIT_GRIPPER1_TYPE: uiOperatorPrompt := UINT#2;
	E_CELL_MANAGER_STATE.WAIT_GRIPPER2_CONTENT: uiOperatorPrompt := UINT#3;
	E_CELL_MANAGER_STATE.WAIT_GRIPPER2_TYPE: uiOperatorPrompt := UINT#4;
	E_CELL_MANAGER_STATE.WAIT_START_MACHINE: uiOperatorPrompt := UINT#5;
ELSE
	uiOperatorPrompt := UINT#0;
END_CASE;
Status.xOperatorPromptActive := uiOperatorPrompt <> UINT#0;
Status.xOperatorChoiceAllowed := Status.xOperatorPromptActive
	AND NOT xManual
	AND NOT xGlobalError
	AND (Error.dwErrorActive = DWORD#0)
	AND xRobotInterfaceReady
	AND xConfigurationValid
	AND xPointsConfigured
	AND xDrivesReady
	AND xRobotReady
	AND xMagazineReady
	AND (NOT xSafetyHomeRequired OR xRobotAtSafetyHome);
Status.xOperatorCancelAllowed := Status.xOperatorPromptActive;
Status.uiOperatorPrompt := uiOperatorPrompt;
Status.uiOperatorTypeMask := uiOperatorTypeMask;
Status.uiOperatorMachineMask := uiOperatorMachineMask;

// Во время TAKE/CHANGE тип будущей заготовки уже известен. Передаём его
// FB_ROBOT до закрытия первого захвата, чтобы авария между CLAMP и DONE не
// оставила физически взятую заготовку с типом 0.
IF ((eMagazineOperation = E_MAGAZINE_OPERATION.TAKE)
	OR (eMagazineOperation = E_MAGAZINE_OPERATION.CHANGE))
AND (uiSelectedType >= UINT#1)
AND (uiSelectedType <= Config.uiTypeCount) THEN
	Command.uiBlankPayloadType := uiSelectedType;
ELSE
	Command.uiBlankPayloadType := uiBlankPayloadType;
END_IF;
Command.uiDetailPayloadType := uiDetailPayloadType;

CASE eState OF
	E_CELL_MANAGER_STATE.IDLE: Diag.eState := E_CELL_STATE.IDLE;
	E_CELL_MANAGER_STATE.PRESTART_IDENTIFY,
	E_CELL_MANAGER_STATE.WAIT_GRIPPER1_CONTENT,
	E_CELL_MANAGER_STATE.WAIT_GRIPPER1_TYPE,
	E_CELL_MANAGER_STATE.WAIT_GRIPPER2_CONTENT,
	E_CELL_MANAGER_STATE.WAIT_GRIPPER2_TYPE,
	E_CELL_MANAGER_STATE.WAIT_START_MACHINE: Diag.eState := E_CELL_STATE.ROUTE_PAYLOAD;
	E_CELL_MANAGER_STATE.PLAN_TARGET, E_CELL_MANAGER_STATE.SELECT_FALLBACK: Diag.eState := E_CELL_STATE.SELECT_MACHINE;
	E_CELL_MANAGER_STATE.MAGAZINE_EXECUTE: Diag.eState := E_CELL_STATE.MAGAZINE;
	E_CELL_MANAGER_STATE.RELEASE_MAGAZINE: Diag.eState := E_CELL_STATE.RELEASE_MAGAZINE;
	E_CELL_MANAGER_STATE.ROUTE_TO_TARGET: Diag.eState := E_CELL_STATE.MOVE_TO_MACHINE;
	E_CELL_MANAGER_STATE.RELEASE_ROBOT_COMMAND: Diag.eState := E_CELL_STATE.RELEASE_ROBOT_COMMAND;
	E_CELL_MANAGER_STATE.WAIT_TARGET: Diag.eState := E_CELL_STATE.WAIT_MACHINE;
	E_CELL_MANAGER_STATE.SERVICE_TARGET: Diag.eState := E_CELL_STATE.SERVICE_MACHINE;
	E_CELL_MANAGER_STATE.MACHINE_FAULT_STOP: Diag.eState := E_CELL_STATE.SERVICE_MACHINE;
	E_CELL_MANAGER_STATE.WAIT_MAGAZINE: Diag.eState := E_CELL_STATE.WAIT_MAGAZINE;
	E_CELL_MANAGER_STATE.GEOMETRY_WAIT_FREE: Diag.eState := E_CELL_STATE.GEOMETRY_WAIT;
	E_CELL_MANAGER_STATE.GEOMETRY_DELIVER, E_CELL_MANAGER_STATE.GEOMETRY_RELEASE_COMMAND: Diag.eState := E_CELL_STATE.GEOMETRY_TRANSFER;
	E_CELL_MANAGER_STATE.TEST_ABORT_STOP: Diag.eState := E_CELL_STATE.IDLE;
	E_CELL_MANAGER_STATE.ERROR: Diag.eState := E_CELL_STATE.ERROR;
END_CASE;

CycleStatus.eState := eState;
CycleStatus.uiSelectedMachine := uiSelectedMachine;
CycleStatus.uiSelectedType := uiSelectedType;
CycleStatus.uiBlankPayloadType := uiBlankPayloadType;
CycleStatus.uiDetailPayloadType := uiDetailPayloadType;
CycleStatus.iTakeSlot := iTakeSlot;
CycleStatus.iPutSlot := iPutSlot;
CycleStatus.xReturningBlank := (eMagazineOperation = E_MAGAZINE_OPERATION.RETURN_BLANK)
	AND ((eState = E_CELL_MANAGER_STATE.MAGAZINE_EXECUTE)
		OR (eState = E_CELL_MANAGER_STATE.RELEASE_MAGAZINE));
CycleStatus.axMachineStartPending := axMachineStartPending;
CycleStatus.auiBlankCount := stMagazineStatus.stTypeStatus.auiBlankCount;
CycleStatus.auiDetailCount := stMagazineStatus.stTypeStatus.auiDetailCount;
CycleStatus.auiFreeCount := stMagazineStatus.stTypeStatus.auiFreeCount;

Error.dwAlarmActive := Error.dwErrorActive;
IF Error.dwErrorActive <> DWORD#0 THEN
	Error.dwErrorLast := Error.dwErrorActive;
END_IF;
Error.stErrorActive := UpdateErrorView(dwError := Error.dwErrorActive);
Error.stErrorLast := UpdateErrorView(dwError := Error.dwErrorLast);
FaultStatus.xResetAllowed := Status.xResetAllowed AND NOT FaultStatus.xBusy;

METHOD PRIVATE IsMachineEligible : BOOL
VAR_INPUT
	uiMachine : UINT; // Проверяемый станок
END_VAR
IsMachineEligible := (uiMachine >= FIRST_MACHINE)
	AND (uiMachine <= LAST_MACHINE);

IF IsMachineEligible THEN
	IsMachineEligible := astMachineStatus[uiMachine].xEnabled
		AND NOT astMachineStatus[uiMachine].xError
		AND NOT astMachineStatus[uiMachine].xDisablePending
		AND NOT axGeometryUnloadBlocked[uiMachine]
		AND (Config.auiMachineType[uiMachine] >= UINT#1)
		AND (Config.auiMachineType[uiMachine] <= Config.uiTypeCount);
END_IF;
END_METHOD

METHOD PRIVATE RaisePayloadRouteWarning
VAR_INPUT
	uiPayloadType     : UINT;
	uiDestinationType : UINT;
END_VAR
IF (uiPayloadType >= UINT#1)
AND (uiDestinationType >= UINT#1)
AND (uiPayloadType <> uiDestinationType) THEN
	IF NOT xPayloadRouteWarningActive THEN
		Diag.stWarning.uiCode := WRN_PAYLOAD_ROUTE_MISMATCH;
		Diag.stWarning.udiSequence := Diag.stWarning.udiSequence + UDINT#1;
		IF Diag.stWarning.udiSequence = UDINT#0 THEN
			Diag.stWarning.udiSequence := UDINT#1;
		END_IF;
		xPayloadRouteWarningActive := TRUE;
	END_IF;
ELSE
	xPayloadRouteWarningActive := FALSE;
END_IF;
END_METHOD

METHOD PRIVATE RunGeometryRoute
CASE eState OF
	E_CELL_MANAGER_STATE.GEOMETRY_WAIT_FREE:
		IF uiGeometryParkStation = UINT#1 THEN eGeometrySafePoint := E_POINT_NAME.GEOMETRY_1_SAFE;
		ELSE eGeometrySafePoint := E_POINT_NAME.GEOMETRY_2_SAFE; END_IF;
		IF stRobotStatus.xBusy OR stRobotStatus.xDone OR xMotionBusy THEN
			// Освобождение ГК не отменяет уже выданное парковочное движение.
			Command.stRobot.xExecute := TRUE; Command.stRobot.eAction := E_ROBOT_ACTION.MOVE_TO_POINT;
			Command.stRobot.eSetPoint := eGeometrySafePoint;
			IF stRobotStatus.xDone THEN eGeometryReturnState := E_CELL_MANAGER_STATE.GEOMETRY_WAIT_FREE; eState := E_CELL_MANAGER_STATE.GEOMETRY_RELEASE_COMMAND; END_IF;
		ELSIF xStopRequested THEN
			xRunning := FALSE; eState := E_CELL_MANAGER_STATE.IDLE;
		ELSIF F_GEOMETRY_SELECT_STATION(xRequireFree := TRUE, uiMachine := uiGeometryMachine) > UINT#0 THEN
			eState := E_CELL_MANAGER_STATE.PLAN_TARGET;
		ELSIF (F_GEOMETRY_SELECT_STATION(xRequireFree := FALSE, uiMachine := uiGeometryMachine) = UINT#0) OR NOT GVL_GEOMETRY_CONTROL.xWaitWhenOccupied THEN
			eState := E_CELL_MANAGER_STATE.PLAN_TARGET;
		ELSE
			// Ожидаем с деталью в захвате на безопасной высоте; конвейер может работать.
			IF uiGeometryParkStation = UINT#1 THEN eGeometrySafePoint := E_POINT_NAME.GEOMETRY_1_SAFE;
			ELSE eGeometrySafePoint := E_POINT_NAME.GEOMETRY_2_SAFE; END_IF;
			IF stRobotStatus.eCurrentPoint <> eGeometrySafePoint THEN
				Command.stRobot.xExecute := TRUE; Command.stRobot.eAction := E_ROBOT_ACTION.MOVE_TO_POINT;
				Command.stRobot.eSetPoint := eGeometrySafePoint;
				IF stRobotStatus.xDone THEN eGeometryReturnState := E_CELL_MANAGER_STATE.GEOMETRY_WAIT_FREE; eState := E_CELL_MANAGER_STATE.GEOMETRY_RELEASE_COMMAND; END_IF;
			END_IF;
		END_IF;
	E_CELL_MANAGER_STATE.GEOMETRY_DELIVER:
		IF (uiGeometryStation < UINT#1) OR (uiGeometryStation > UINT#2) THEN
			Error.dwErrorActive := Error.dwErrorActive OR ERR_ROBOT; eState := E_CELL_MANAGER_STATE.ERROR;
		ELSIF GVL_GEOMETRY_CONTROL.astStatus[uiGeometryStation].xError
		AND NOT GVL_GEOMETRY_CONTROL.astSignals[uiGeometryStation].xRobotInteraction THEN
			// Оборудование отказало до входа: робот может выбрать другой ГК.
			GVL_GEOMETRY_CONTROL.astSignals[uiGeometryStation].xReserve := FALSE;
			GVL_GEOMETRY_CONTROL.astSignals[uiGeometryStation].xReleased := TRUE;
			GVL_GEOMETRY_CONTROL.astCalls[uiGeometryMachine].uiStation := UINT#0;
			GVL_GEOMETRY_CONTROL.astCalls[uiGeometryMachine].uiState := UINT#2;
			GVL_GEOMETRY_CONTROL.astCalls[uiGeometryMachine].uiReason := UINT#4;
			F_GEOMETRY_EVENT(Call := GVL_GEOMETRY_CONTROL.astCalls[uiGeometryMachine]);
			uiGeometryStation := UINT#0; eState := E_CELL_MANAGER_STATE.PLAN_TARGET;
		ELSIF NOT GVL_GEOMETRY_CONTROL.astSignals[uiGeometryStation].xRobotInteraction
		AND (NOT GVL_GEOMETRY_CONTROL.astStatus[uiGeometryStation].xEnabled
			OR (GVL_GEOMETRY_CONTROL.astStatus[uiGeometryStation].uiState = UINT#5)
			OR GVL_GEOMETRY_CONTROL.astStatus[uiGeometryStation].xDriveRunning) THEN
			// Выключение в том же скане, что резерв, не разрешает вход робота.
			GVL_GEOMETRY_CONTROL.astSignals[uiGeometryStation].xReserve := FALSE;
			GVL_GEOMETRY_CONTROL.astSignals[uiGeometryStation].xReleased := TRUE;
			GVL_GEOMETRY_CONTROL.astCalls[uiGeometryMachine].uiStation := UINT#0;
			GVL_GEOMETRY_CONTROL.astCalls[uiGeometryMachine].uiState := UINT#2;
			GVL_GEOMETRY_CONTROL.astCalls[uiGeometryMachine].uiReason := UINT#3;
			F_GEOMETRY_EVENT(Call := GVL_GEOMETRY_CONTROL.astCalls[uiGeometryMachine]);
			uiGeometryStation := UINT#0; eState := E_CELL_MANAGER_STATE.PLAN_TARGET;
		ELSIF GVL_GEOMETRY_CONTROL.astStatus[uiGeometryStation].xError OR stRobotStatus.xError OR xGlobalError THEN
			xSafetyHomeRequired := TRUE; xStoppedPoseValid := FALSE;
			Error.dwErrorActive := Error.dwErrorActive OR ERR_ROBOT; eState := E_CELL_MANAGER_STATE.ERROR;
		ELSIF GVL_GEOMETRY_CONTROL.astStatus[uiGeometryStation].xReserved THEN
			IF uiGeometryStation = UINT#1 THEN
				eGeometrySafePoint := E_POINT_NAME.GEOMETRY_1_SAFE; eGeometryPlacePoint := E_POINT_NAME.GEOMETRY_1_PLACE;
			ELSE
				eGeometrySafePoint := E_POINT_NAME.GEOMETRY_2_SAFE; eGeometryPlacePoint := E_POINT_NAME.GEOMETRY_2_PLACE;
			END_IF;
			GVL_GEOMETRY_CONTROL.astSignals[uiGeometryStation].xRobotInteraction := TRUE;
			IF uiGeometryStep <= UINT#4 THEN
				Command.stRobot.xExecute := TRUE; Command.stRobot.eAction := E_ROBOT_ACTION.MOVE_TO_POINT;
				CASE uiGeometryStep OF
					UINT#0, UINT#4: Command.stRobot.eSetPoint := eGeometrySafePoint;
					// Для укладки на ГК нужна ориентация «к заготовке»; поворот выполняется на SAFE.
					UINT#1: Command.stRobot.eAction := E_ROBOT_ACTION.ROTATE_TO_BLANK;
					UINT#2: Command.stRobot.eSetPoint := eGeometryPlacePoint;
					UINT#3: Command.stRobot.eAction := E_ROBOT_ACTION.UNCLAMP_2;
				END_CASE;
				IF stRobotStatus.xDone THEN
					IF uiGeometryStep = UINT#3 THEN
						IF stRobotStatus.xGripper2Open AND NOT stRobotStatus.xDetailAvailable THEN
							GVL_GEOMETRY_CONTROL.astSignals[uiGeometryStation].xDeposited := TRUE;
							uiDetailPayloadType := UINT#0;
						ELSE Error.dwErrorActive := Error.dwErrorActive OR ERR_ROBOT; eState := E_CELL_MANAGER_STATE.ERROR; END_IF;
					END_IF;
					IF eState <> E_CELL_MANAGER_STATE.ERROR THEN
						eGeometryReturnState := E_CELL_MANAGER_STATE.GEOMETRY_DELIVER;
						eState := E_CELL_MANAGER_STATE.GEOMETRY_RELEASE_COMMAND;
					END_IF;
				END_IF;
			ELSE
				GVL_GEOMETRY_CONTROL.astSignals[uiGeometryStation].xReserve := FALSE;
				GVL_GEOMETRY_CONTROL.astSignals[uiGeometryStation].xDeposited := FALSE;
				GVL_GEOMETRY_CONTROL.astSignals[uiGeometryStation].xRobotInteraction := FALSE;
				GVL_GEOMETRY_CONTROL.astSignals[uiGeometryStation].xReleased := TRUE;
				GVL_GEOMETRY_CONTROL.uiLastStation := uiGeometryStation;
				xGeometryHeld := FALSE; uiGeometryMachine := UINT#0; uiGeometryStation := UINT#0;
				eState := E_CELL_MANAGER_STATE.PLAN_TARGET;
			END_IF;
		ELSE
			// Потеря резерва в зоне робота требует восстановления, а не нового маршрута.
			IF GVL_GEOMETRY_CONTROL.astSignals[uiGeometryStation].xRobotInteraction THEN
				xSafetyHomeRequired := TRUE; xStoppedPoseValid := FALSE;
				Error.dwErrorActive := Error.dwErrorActive OR ERR_ROBOT; eState := E_CELL_MANAGER_STATE.ERROR;
			ELSIF NOT GVL_GEOMETRY_CONTROL.astStatus[uiGeometryStation].xReady
			OR (GVL_GEOMETRY_CONTROL.astStatus[uiGeometryStation].uiState = UINT#5) THEN
				GVL_GEOMETRY_CONTROL.astSignals[uiGeometryStation].xReserve := FALSE;
				GVL_GEOMETRY_CONTROL.astSignals[uiGeometryStation].xReleased := TRUE;
				GVL_GEOMETRY_CONTROL.astCalls[uiGeometryMachine].uiStation := UINT#0;
				GVL_GEOMETRY_CONTROL.astCalls[uiGeometryMachine].uiState := UINT#2;
				GVL_GEOMETRY_CONTROL.astCalls[uiGeometryMachine].uiReason := UINT#3;
				F_GEOMETRY_EVENT(Call := GVL_GEOMETRY_CONTROL.astCalls[uiGeometryMachine]);
				uiGeometryStation := UINT#0; eState := E_CELL_MANAGER_STATE.PLAN_TARGET;
			END_IF;
		END_IF;
	E_CELL_MANAGER_STATE.GEOMETRY_RELEASE_COMMAND:
		IF stRobotStatus.xError THEN
			xSafetyHomeRequired := TRUE; xStoppedPoseValid := FALSE;
			Error.dwErrorActive := Error.dwErrorActive OR ERR_ROBOT; eState := E_CELL_MANAGER_STATE.ERROR;
		ELSIF NOT stRobotStatus.xBusy AND NOT stRobotStatus.xDone THEN
			IF eGeometryReturnState = E_CELL_MANAGER_STATE.GEOMETRY_DELIVER THEN uiGeometryStep := uiGeometryStep + UINT#1; END_IF;
			eState := eGeometryReturnState;
		END_IF;
END_CASE;
END_METHOD

METHOD PRIVATE IsMachineCompatible : BOOL
VAR_INPUT
	uiMachine     : UINT; // Проверяемый станок
	uiProductType : UINT; // Тип заготовки в захвате
END_VAR
IsMachineCompatible := IsMachineEligible(uiMachine := uiMachine);
IF IsMachineCompatible THEN
	IsMachineCompatible := (uiProductType >= UINT#1)
		AND (uiProductType <= Config.uiTypeCount)
		AND (Config.auiMachineType[uiMachine] = uiProductType);
END_IF;
END_METHOD

METHOD PRIVATE SelectMachineBeforeTake : UINT
VAR
	uiMachine           : UINT; // Проверяемый станок
	uiType              : UINT; // Тип станка
	xTimedFound         : BOOL; // Найден кандидат с оценкой времени
	tMinimumRemaining   : TIME; // Минимальное найденное оставшееся время
	tCandidateRemaining : TIME; // Оценка кандидата, который подтверждает запуск цикла
END_VAR
SelectMachineBeforeTake := UINT#0;
xTimedFound := FALSE;
tMinimumRemaining := T#0S;

// Сначала выбирается станок, который можно обслужить без ожидания.
// xPartReady отдельно не используется: после завершения обслуживания он может
// сохраняться до перехода FB_MACHINE из DONE в IDLE и повторно выбрать тот же станок.
FOR uiMachine := FIRST_MACHINE TO LAST_MACHINE DO
	uiType := Config.auiMachineType[uiMachine];
	IF IsMachineEligible(uiMachine := uiMachine) THEN
		IF (SelectMachineBeforeTake = UINT#0)
		AND (stMagazineStatus.stTypeStatus.aiBlankSlot[uiType] > SINT#0)
		AND astMachineStatus[uiMachine].xCanAcceptService
		AND ((astMachineStatus[uiMachine].ePartState = E_PART_STATE.EMPTY)
			OR astMachineStatus[uiMachine].xServiceRequired) THEN
			SelectMachineBeforeTake := uiMachine;
		END_IF;
	END_IF;
END_FOR;

// Затем сравниваются фактически обрабатывающие станки по оставшемуся времени.
IF SelectMachineBeforeTake = UINT#0 THEN
	FOR uiMachine := FIRST_MACHINE TO LAST_MACHINE DO
		uiType := Config.auiMachineType[uiMachine];
		IF IsMachineEligible(uiMachine := uiMachine) THEN
			IF (stMagazineStatus.stTypeStatus.aiBlankSlot[uiType] > SINT#0)
			AND astMachineStatus[uiMachine].xProcessing
			AND astMachineStatus[uiMachine].xCycleTimeValid THEN
				IF NOT xTimedFound
				OR (astMachineStatus[uiMachine].tRemaining < tMinimumRemaining) THEN
					SelectMachineBeforeTake := uiMachine;
					tMinimumRemaining := astMachineStatus[uiMachine].tRemaining;
					xTimedFound := TRUE;
				END_IF;
			END_IF;
		END_IF;
	END_FOR;
END_IF;

// Только что обслуженный станок может появиться в xProcessing на несколько циклов PLC позже.
// До подтверждения запуска он участвует в том же сравнении по полному tCycleExpected.
IF (SelectMachineBeforeTake = UINT#0) OR xTimedFound THEN
	FOR uiMachine := FIRST_MACHINE TO LAST_MACHINE DO
		uiType := Config.auiMachineType[uiMachine];
		IF axMachineStartPending[uiMachine]
		AND IsMachineEligible(uiMachine := uiMachine)
		AND (stMagazineStatus.stTypeStatus.aiBlankSlot[uiType] > SINT#0)
		AND astMachineStatus[uiMachine].xCycleTimeValid THEN
			tCandidateRemaining := START_PENDING_ESTIMATE
				+ astMachineStatus[uiMachine].tCycleExpected;
			IF NOT xTimedFound
			OR (tCandidateRemaining < tMinimumRemaining) THEN
				SelectMachineBeforeTake := uiMachine;
				tMinimumRemaining := tCandidateRemaining;
				xTimedFound := TRUE;
			END_IF;
		END_IF;
	END_FOR;
END_IF;

// Неизвестное время не делает включённый исправный станок недоступным.
IF (SelectMachineBeforeTake = UINT#0) AND NOT xTimedFound THEN
	FOR uiMachine := FIRST_MACHINE TO LAST_MACHINE DO
		uiType := Config.auiMachineType[uiMachine];
		IF IsMachineEligible(uiMachine := uiMachine) THEN
			IF (SelectMachineBeforeTake = UINT#0)
			AND (stMagazineStatus.stTypeStatus.aiBlankSlot[uiType] > SINT#0)
			AND (astMachineStatus[uiMachine].xProcessing
				OR axMachineStartPending[uiMachine]) THEN
				SelectMachineBeforeTake := uiMachine;
			END_IF;
		END_IF;
	END_FOR;
END_IF;
END_METHOD

METHOD PRIVATE PlanGeometry : BOOL
VAR
	uiFree : UINT;
	uiAvailable : UINT;
END_VAR
PlanGeometry := FALSE;
IF xGeometryHeld AND stRobotStatus.xDetailAvailable AND (uiGeometryMachine >= UINT#1) AND (uiGeometryMachine <= UINT#3) THEN
	uiFree := F_GEOMETRY_SELECT_STATION(xRequireFree := TRUE, uiMachine := uiGeometryMachine);
	uiAvailable := F_GEOMETRY_SELECT_STATION(xRequireFree := FALSE, uiMachine := uiGeometryMachine);
	IF uiFree > UINT#0 THEN
		uiGeometryStation := uiFree; uiGeometryStep := UINT#0;
		GVL_GEOMETRY_CONTROL.astCalls[uiGeometryMachine].uiStation := uiFree;
		GVL_GEOMETRY_CONTROL.astCalls[uiGeometryMachine].uiState := UINT#3;
		GVL_GEOMETRY_CONTROL.astCalls[uiGeometryMachine].uiReason := UINT#0;
		F_GEOMETRY_EVENT(Call := GVL_GEOMETRY_CONTROL.astCalls[uiGeometryMachine]);
		GVL_GEOMETRY_CONTROL.astSignals[uiFree].Call := GVL_GEOMETRY_CONTROL.astCalls[uiGeometryMachine];
		GVL_GEOMETRY_CONTROL.astSignals[uiFree].xReserve := TRUE;
		eState := E_CELL_MANAGER_STATE.GEOMETRY_DELIVER; PlanGeometry := TRUE;
	ELSIF (uiAvailable > UINT#0) AND GVL_GEOMETRY_CONTROL.xWaitWhenOccupied THEN
		uiGeometryParkStation := uiAvailable;
		eState := E_CELL_MANAGER_STATE.GEOMETRY_WAIT_FREE; PlanGeometry := TRUE;
	ELSE
		// Окончательный журнал магазина формируем только по фактической укладке.
		IF uiAvailable > UINT#0 THEN uiGeometryBypassReason := UINT#1; ELSE uiGeometryBypassReason := UINT#2; END_IF;
		udiGeometryMagazineCounter := stMagazineStatus.udiProducedPartsTotal;
	END_IF;
END_IF;
END_METHOD

METHOD PRIVATE UpdateErrorView : ST_CELL_ERROR
VAR_INPUT
	dwError : DWORD; // Битовая маска ошибок нового менеджера
END_VAR
VAR
	stError : ST_CELL_ERROR; // Совместимое представление ошибок
END_VAR
stError.BOTH_GRIPPERS_OCCUPIED := (dwError AND ERR_BOTH_GRIPPERS) <> DWORD#0;
stError.ROBOT_ERROR := (dwError AND ERR_ROBOT) <> DWORD#0;
stError.MAGAZINE_ERROR := (dwError AND ERR_MAGAZINE) <> DWORD#0;
stError.MACHINE_ERROR := (dwError AND ERR_MACHINE) <> DWORD#0;
stError.GLOBAL_STOP := (dwError AND ERR_GLOBAL_STOP) <> DWORD#0;
UpdateErrorView := stError;
END_METHOD

METHOD PRIVATE SelectMachineForUnload : UINT
VAR_INPUT
	uiCurrentMachine : UINT; // Текущая цель для устойчивого повторного выбора
END_VAR
VAR
	uiMachine           : UINT; // Проверяемый станок
	uiType              : UINT; // Тип детали станка
	xTimedFound         : BOOL; // Найден станок с оценкой времени
	xCurrentTimed       : BOOL; // Текущая цель имеет сопоставимую оценку
	tMinimumRemaining   : TIME; // Минимальное найденное оставшееся время
	tCandidateRemaining : TIME; // Оценка проверяемого станка
	tCurrentRemaining   : TIME; // Оценка текущей цели
END_VAR
SelectMachineForUnload := UINT#0;
xTimedFound := FALSE;
xCurrentTimed := FALSE;
tMinimumRemaining := T#0S;
tCandidateRemaining := T#0S;
tCurrentRemaining := T#0S;

// Если робот уже ждёт над готовым станком, лишнее перемещение не требуется.
IF (uiCurrentMachine >= FIRST_MACHINE)
AND (uiCurrentMachine <= LAST_MACHINE) THEN
	IF IsMachineEligible(uiMachine := uiCurrentMachine) THEN
		uiType := Config.auiMachineType[uiCurrentMachine];
		IF (stMagazineStatus.stTypeStatus.aiFreeSlot[uiType] > SINT#0)
		AND astMachineStatus[uiCurrentMachine].xCanAcceptService
		AND astMachineStatus[uiCurrentMachine].xServiceRequired
		AND (astMachineStatus[uiCurrentMachine].ePartState = E_PART_STATE.LOADED)
		AND (astMachineStatus[uiCurrentMachine].ePartType = E_PART_TYPE.DETAIL) THEN
			SelectMachineForUnload := uiCurrentMachine;
		END_IF;
	END_IF;
END_IF;

// Готовая деталь имеет приоритет над ожиданием обработки.
FOR uiMachine := FIRST_MACHINE TO LAST_MACHINE DO
	uiType := Config.auiMachineType[uiMachine];
	IF IsMachineEligible(uiMachine := uiMachine) THEN
		IF (SelectMachineForUnload = UINT#0)
		AND astMachineStatus[uiMachine].xCanAcceptService
		AND astMachineStatus[uiMachine].xServiceRequired
		AND (astMachineStatus[uiMachine].ePartState = E_PART_STATE.LOADED)
		AND (astMachineStatus[uiMachine].ePartType = E_PART_TYPE.DETAIL)
		AND (stMagazineStatus.stTypeStatus.aiFreeSlot[uiType] > SINT#0) THEN
			SelectMachineForUnload := uiMachine;
		END_IF;
	END_IF;
END_FOR;

// Если готовых деталей пока нет, робот заранее направляется к станку с
// минимальным оставшимся временем обработки.
IF SelectMachineForUnload = UINT#0 THEN
	FOR uiMachine := FIRST_MACHINE TO LAST_MACHINE DO
		uiType := Config.auiMachineType[uiMachine];
		IF IsMachineEligible(uiMachine := uiMachine) THEN
			IF (stMagazineStatus.stTypeStatus.aiFreeSlot[uiType] > SINT#0)
			AND astMachineStatus[uiMachine].xCycleTimeValid THEN
				IF astMachineStatus[uiMachine].xProcessing THEN
					tCandidateRemaining := astMachineStatus[uiMachine].tRemaining;
				ELSIF axMachineStartPending[uiMachine] THEN
					tCandidateRemaining := START_PENDING_ESTIMATE
						+ astMachineStatus[uiMachine].tCycleExpected;
				ELSE
					tCandidateRemaining := T#0S;
				END_IF;

				IF astMachineStatus[uiMachine].xProcessing
				OR axMachineStartPending[uiMachine] THEN
					IF NOT xTimedFound
					OR (tCandidateRemaining < tMinimumRemaining) THEN
						SelectMachineForUnload := uiMachine;
						tMinimumRemaining := tCandidateRemaining;
						xTimedFound := TRUE;
					END_IF;
				END_IF;
			END_IF;
		END_IF;
	END_FOR;

	// При почти одинаковом времени сохраняется уже выбранная цель.
	IF xTimedFound
	AND (uiCurrentMachine >= FIRST_MACHINE)
	AND (uiCurrentMachine <= LAST_MACHINE) THEN
		IF (SelectMachineForUnload <> uiCurrentMachine)
		AND IsMachineEligible(uiMachine := uiCurrentMachine) THEN
			uiType := Config.auiMachineType[uiCurrentMachine];
			IF (stMagazineStatus.stTypeStatus.aiFreeSlot[uiType] > SINT#0)
			AND astMachineStatus[uiCurrentMachine].xCycleTimeValid THEN
				xCurrentTimed := astMachineStatus[uiCurrentMachine].xProcessing
					OR axMachineStartPending[uiCurrentMachine];
				IF astMachineStatus[uiCurrentMachine].xProcessing THEN
					tCurrentRemaining := astMachineStatus[uiCurrentMachine].tRemaining;
				ELSIF axMachineStartPending[uiCurrentMachine] THEN
					tCurrentRemaining := START_PENDING_ESTIMATE
						+ astMachineStatus[uiCurrentMachine].tCycleExpected;
				END_IF;
				IF xCurrentTimed
				AND (tCurrentRemaining >= tMinimumRemaining)
				AND ((tCurrentRemaining - tMinimumRemaining) <= MACHINE_SWITCH_DEADBAND) THEN
					SelectMachineForUnload := uiCurrentMachine;
				END_IF;
			END_IF;
		END_IF;
	END_IF;
END_IF;

// При неизвестном времени сохраняется текущая цель либо выбирается первый
// обрабатывающийся/только что запущенный станок с доступным слотом.
IF SelectMachineForUnload = UINT#0 THEN
	IF (uiCurrentMachine >= FIRST_MACHINE)
	AND (uiCurrentMachine <= LAST_MACHINE) THEN
		IF IsMachineEligible(uiMachine := uiCurrentMachine) THEN
			uiType := Config.auiMachineType[uiCurrentMachine];
			IF (stMagazineStatus.stTypeStatus.aiFreeSlot[uiType] > SINT#0)
			AND (astMachineStatus[uiCurrentMachine].xProcessing
				OR axMachineStartPending[uiCurrentMachine]) THEN
				SelectMachineForUnload := uiCurrentMachine;
			END_IF;
		END_IF;
	END_IF;

	FOR uiMachine := FIRST_MACHINE TO LAST_MACHINE DO
		uiType := Config.auiMachineType[uiMachine];
		IF IsMachineEligible(uiMachine := uiMachine) THEN
			IF (SelectMachineForUnload = UINT#0)
			AND (stMagazineStatus.stTypeStatus.aiFreeSlot[uiType] > SINT#0)
			AND (astMachineStatus[uiMachine].xProcessing
				OR axMachineStartPending[uiMachine]) THEN
				SelectMachineForUnload := uiMachine;
			END_IF;
		END_IF;
	END_FOR;
END_IF;

// Переход от окончания цикла к готовности двери может занять несколько сканов.
// В это время сохраняется станок с физически загруженной деталью/заготовкой.
IF SelectMachineForUnload = UINT#0 THEN
	IF (uiCurrentMachine >= FIRST_MACHINE)
	AND (uiCurrentMachine <= LAST_MACHINE) THEN
		IF IsMachineEligible(uiMachine := uiCurrentMachine) THEN
			uiType := Config.auiMachineType[uiCurrentMachine];
			IF (stMagazineStatus.stTypeStatus.aiFreeSlot[uiType] > SINT#0)
			AND (astMachineStatus[uiCurrentMachine].ePartState = E_PART_STATE.LOADED)
			AND ((astMachineStatus[uiCurrentMachine].ePartType = E_PART_TYPE.PART)
				OR (astMachineStatus[uiCurrentMachine].ePartType = E_PART_TYPE.DETAIL)) THEN
				SelectMachineForUnload := uiCurrentMachine;
			END_IF;
		END_IF;
	END_IF;

	FOR uiMachine := FIRST_MACHINE TO LAST_MACHINE DO
		uiType := Config.auiMachineType[uiMachine];
		IF IsMachineEligible(uiMachine := uiMachine) THEN
			IF (SelectMachineForUnload = UINT#0)
			AND (stMagazineStatus.stTypeStatus.aiFreeSlot[uiType] > SINT#0)
			AND (astMachineStatus[uiMachine].ePartState = E_PART_STATE.LOADED)
			AND ((astMachineStatus[uiMachine].ePartType = E_PART_TYPE.PART)
				OR (astMachineStatus[uiMachine].ePartType = E_PART_TYPE.DETAIL)) THEN
				SelectMachineForUnload := uiMachine;
			END_IF;
		END_IF;
	END_FOR;
END_IF;
END_METHOD

METHOD PRIVATE UpdateGeometryWait
VAR
	uiMachine : UINT;
	uiFreeStation : UINT;
	uiFirstCallMachine : UINT;
	uiCallState : UINT;
	xCalled : BOOL;
	xReadyDetail : BOOL;
	xWaiting : BOOL;
	xRaiseWarning : BOOL;
	Call : ST_GEOMETRY_CALL;
	EmptyCall : ST_GEOMETRY_CALL;
END_VAR
uiFreeStation := F_GEOMETRY_SELECT_STATION(xRequireFree := TRUE, uiMachine := UINT#0);
xRaiseWarning := FALSE;
FOR uiMachine := FIRST_MACHINE TO LAST_MACHINE DO
	uiCallState := GVL_GEOMETRY_CONTROL.astCalls[uiMachine].uiState;
	xCalled := uiCallState = UINT#1;
	// Автовызов известен до выгрузки; счётчик меняется только при фактическом взятии.
	IF ((uiCallState = UINT#0) OR (uiCallState > UINT#3))
	AND GVL_GEOMETRY_CONTROL.xSupported AND GVL_GEOMETRY_CONTROL.xAutoEnabled
	AND (GVL_GEOMETRY_CONTROL.astStatus[1].xEnabled OR GVL_GEOMETRY_CONTROL.astStatus[2].xEnabled)
	AND (GVL_GEOMETRY_CONTROL.auiActiveCount[uiMachine] >= (MAX(UINT#1, GVL_GEOMETRY_CONTROL.auiPeriod[uiMachine]) - UINT#1)) THEN
		xCalled := TRUE;
	END_IF;
	xReadyDetail := astMachineStatus[uiMachine].xEnabled
		AND NOT astMachineStatus[uiMachine].xError AND NOT astMachineStatus[uiMachine].xDisablePending
		AND NOT astMachineStatus[uiMachine].xBusy AND NOT astMachineStatus[uiMachine].xProcessing
		AND astMachineStatus[uiMachine].xCanAcceptService AND astMachineStatus[uiMachine].xServiceRequired
		AND (astMachineStatus[uiMachine].ePartState = E_PART_STATE.LOADED)
		AND (astMachineStatus[uiMachine].ePartType = E_PART_TYPE.DETAIL);
	IF xRunning AND NOT xManual AND xCalled AND xReadyDetail AND (uiCallState <> UINT#1) THEN
		GVL_GEOMETRY_CONTROL.udiNextCallId := GVL_GEOMETRY_CONTROL.udiNextCallId + UDINT#1;
		IF GVL_GEOMETRY_CONTROL.udiNextCallId = UDINT#0 THEN GVL_GEOMETRY_CONTROL.udiNextCallId := UDINT#1; END_IF;
		Call := EmptyCall; Call.udiId := GVL_GEOMETRY_CONTROL.udiNextCallId;
		Call.uiMachine := uiMachine; Call.uiProductType := Config.auiMachineType[uiMachine]; Call.uiState := UINT#1;
		GVL_GEOMETRY_CONTROL.astCalls[uiMachine] := Call;
		F_GEOMETRY_EVENT(Call := Call);
	END_IF;
	// Пустой станок можно загрузить. Уже начатый рецепт не прерываем.
	axGeometryUnloadBlocked[uiMachine] := xCalled AND (uiFreeStation = UINT#0)
		AND (astMachineStatus[uiMachine].ePartState = E_PART_STATE.LOADED)
		AND NOT astMachineStatus[uiMachine].xBusy;
END_FOR;

// Выбираем голову после создания всех автовызовов этого скана.
uiFirstCallMachine := F_GEOMETRY_FIRST_CALL();
FOR uiMachine := FIRST_MACHINE TO LAST_MACHINE DO
	IF (GVL_GEOMETRY_CONTROL.astCalls[uiMachine].uiState = UINT#1)
	AND (uiMachine <> uiFirstCallMachine)
	AND (astMachineStatus[uiMachine].ePartState = E_PART_STATE.LOADED)
	AND NOT astMachineStatus[uiMachine].xBusy THEN
		// Более поздний вызов не обгоняет первый, даже если его деталь уже готова.
		axGeometryUnloadBlocked[uiMachine] := TRUE;
	END_IF;
	xReadyDetail := astMachineStatus[uiMachine].xEnabled
		AND NOT astMachineStatus[uiMachine].xError AND NOT astMachineStatus[uiMachine].xDisablePending
		AND NOT astMachineStatus[uiMachine].xBusy AND NOT astMachineStatus[uiMachine].xProcessing
		AND astMachineStatus[uiMachine].xCanAcceptService AND astMachineStatus[uiMachine].xServiceRequired
		AND (astMachineStatus[uiMachine].ePartState = E_PART_STATE.LOADED)
		AND (astMachineStatus[uiMachine].ePartType = E_PART_TYPE.DETAIL);
	// Ожидание своей очереди при свободном ГК не является причиной W52.
	xWaiting := xRunning AND NOT xManual AND NOT xGlobalError
		AND xReadyDetail AND axGeometryUnloadBlocked[uiMachine] AND (uiFreeStation = UINT#0);
	// Отдельный TON для каждого вызова; реальное время, без ускорения симуляции.
	atonGeometryWait[uiMachine](IN := xWaiting AND NOT GVL_ALARM.Command.xResetWarnings
		AND (audiGeometryWaitCallId[uiMachine] = GVL_GEOMETRY_CONTROL.astCalls[uiMachine].udiId),
		PT := GVL_GEOMETRY_CONTROL.tWaitWarningTimeout);
	IF NOT xWaiting OR GVL_ALARM.Command.xResetWarnings
	OR (audiGeometryWaitCallId[uiMachine] <> GVL_GEOMETRY_CONTROL.astCalls[uiMachine].udiId) THEN
		axGeometryWaitWarned[uiMachine] := FALSE;
	END_IF;
	audiGeometryWaitCallId[uiMachine] := GVL_GEOMETRY_CONTROL.astCalls[uiMachine].udiId;
	IF atonGeometryWait[uiMachine].Q AND NOT axGeometryWaitWarned[uiMachine] THEN
		axGeometryWaitWarned[uiMachine] := TRUE; xRaiseWarning := TRUE;
	END_IF;
END_FOR;
IF xRaiseWarning THEN
	GVL_GEOMETRY_CONTROL.stCellWarning.uiCode := WRN_GEOMETRY_WAIT_TIMEOUT; // WARNING: остальные станки продолжают работу
	GVL_GEOMETRY_CONTROL.stCellWarning.udiSequence := GVL_GEOMETRY_CONTROL.stCellWarning.udiSequence + UDINT#1;
	IF GVL_GEOMETRY_CONTROL.stCellWarning.udiSequence = UDINT#0 THEN GVL_GEOMETRY_CONTROL.stCellWarning.udiSequence := UDINT#1; END_IF;
END_IF;
END_METHOD

METHOD PRIVATE SelectMachineForHeldBlank : UINT
VAR_INPUT
	uiProductType    : UINT; // Тип уже взятой заготовки
	uiCurrentMachine : UINT; // Текущая цель для устойчивого повторного выбора
END_VAR
VAR
	uiMachine           : UINT; // Проверяемый станок
	xTimedFound         : BOOL; // Найден станок с оценкой времени
	xCurrentTimed       : BOOL; // Текущая цель имеет сопоставимую оценку
	tMinimumRemaining   : TIME; // Минимальное оставшееся время
	tCandidateRemaining : TIME; // Оценка проверяемого станка
	tCurrentRemaining   : TIME; // Оценка текущей цели
END_VAR
SelectMachineForHeldBlank := UINT#0;
xTimedFound := FALSE;
xCurrentTimed := FALSE;
tMinimumRemaining := T#0S;
tCandidateRemaining := T#0S;
tCurrentRemaining := T#0S;

// UINT#0 означает, что после остановки/аварии текущая цель ещё не выбрана.
// Проверка диапазона вынесена отдельно: обычный AND в CODESYS вычисляет все
// операнды и не защищает ARRAY [1..3] от обращения по индексу 0.
IF (uiCurrentMachine >= FIRST_MACHINE)
AND (uiCurrentMachine <= LAST_MACHINE) THEN
	// Если робот уже находится у готовой совместимой цели, лишнее перемещение не требуется.
	IF IsMachineCompatible(
		uiMachine := uiCurrentMachine,
		uiProductType := uiProductType
	)
	AND astMachineStatus[uiCurrentMachine].xCanAcceptService
	AND ((astMachineStatus[uiCurrentMachine].ePartState = E_PART_STATE.EMPTY)
		OR astMachineStatus[uiCurrentMachine].xServiceRequired) THEN
		SelectMachineForHeldBlank := uiCurrentMachine;
	END_IF;
END_IF;

// Готовая совместимая цель имеет приоритет. Переходный xPartReady без
// xCanAcceptService не считается разрешением на повторное обслуживание.
FOR uiMachine := FIRST_MACHINE TO LAST_MACHINE DO
	IF (SelectMachineForHeldBlank = UINT#0)
	AND IsMachineEligible(uiMachine := uiMachine)
	AND (Config.auiMachineType[uiMachine] = uiProductType)
	AND astMachineStatus[uiMachine].xCanAcceptService
	AND ((astMachineStatus[uiMachine].ePartState = E_PART_STATE.EMPTY)
		OR astMachineStatus[uiMachine].xServiceRequired) THEN
		SelectMachineForHeldBlank := uiMachine;
	END_IF;
END_FOR;

// Обрабатывающие и только что запущенные совместимые станки сравниваются
// по одному прогнозу: tRemaining либо полный tCycleExpected для start-pending.
IF SelectMachineForHeldBlank = UINT#0 THEN
	FOR uiMachine := FIRST_MACHINE TO LAST_MACHINE DO
		IF IsMachineEligible(uiMachine := uiMachine)
		AND (Config.auiMachineType[uiMachine] = uiProductType)
		AND astMachineStatus[uiMachine].xCycleTimeValid THEN
			IF astMachineStatus[uiMachine].xProcessing THEN
				tCandidateRemaining := astMachineStatus[uiMachine].tRemaining;
			ELSIF axMachineStartPending[uiMachine] THEN
				tCandidateRemaining := START_PENDING_ESTIMATE
					+ astMachineStatus[uiMachine].tCycleExpected;
			ELSE
				tCandidateRemaining := T#0S;
			END_IF;

			IF astMachineStatus[uiMachine].xProcessing
			OR axMachineStartPending[uiMachine] THEN
				IF NOT xTimedFound
				OR (tCandidateRemaining < tMinimumRemaining) THEN
					SelectMachineForHeldBlank := uiMachine;
					tMinimumRemaining := tCandidateRemaining;
					xTimedFound := TRUE;
				END_IF;
			END_IF;
		END_IF;
	END_FOR;

	// При почти одинаковом времени сохраняется текущая цель.
	IF xTimedFound
	AND (uiCurrentMachine >= FIRST_MACHINE)
	AND (uiCurrentMachine <= LAST_MACHINE) THEN
		IF (SelectMachineForHeldBlank <> uiCurrentMachine)
		AND IsMachineCompatible(
			uiMachine := uiCurrentMachine,
			uiProductType := uiProductType
		)
		AND astMachineStatus[uiCurrentMachine].xCycleTimeValid THEN
			xCurrentTimed := astMachineStatus[uiCurrentMachine].xProcessing
				OR axMachineStartPending[uiCurrentMachine];
			IF astMachineStatus[uiCurrentMachine].xProcessing THEN
				tCurrentRemaining := astMachineStatus[uiCurrentMachine].tRemaining;
			ELSIF axMachineStartPending[uiCurrentMachine] THEN
				tCurrentRemaining := START_PENDING_ESTIMATE
					+ astMachineStatus[uiCurrentMachine].tCycleExpected;
			END_IF;
			IF xCurrentTimed
			AND (tCurrentRemaining >= tMinimumRemaining)
			AND ((tCurrentRemaining - tMinimumRemaining) <= MACHINE_SWITCH_DEADBAND) THEN
				SelectMachineForHeldBlank := uiCurrentMachine;
			END_IF;
		END_IF;
	END_IF;
END_IF;

// Без точной оценки сохраняется текущий обрабатывающий маршрут либо выбирается
// первый совместимый обрабатывающий/start-pending станок.
IF SelectMachineForHeldBlank = UINT#0 THEN
	IF (uiCurrentMachine >= FIRST_MACHINE)
	AND (uiCurrentMachine <= LAST_MACHINE) THEN
		IF IsMachineCompatible(
			uiMachine := uiCurrentMachine,
			uiProductType := uiProductType
		)
		AND (astMachineStatus[uiCurrentMachine].xProcessing
			OR axMachineStartPending[uiCurrentMachine]) THEN
			SelectMachineForHeldBlank := uiCurrentMachine;
		END_IF;
	END_IF;

	FOR uiMachine := FIRST_MACHINE TO LAST_MACHINE DO
		IF (SelectMachineForHeldBlank = UINT#0)
		AND IsMachineEligible(uiMachine := uiMachine)
		AND (Config.auiMachineType[uiMachine] = uiProductType)
		AND (astMachineStatus[uiMachine].xProcessing
			OR axMachineStartPending[uiMachine]) THEN
			SelectMachineForHeldBlank := uiMachine;
		END_IF;
	END_FOR;
END_IF;

// Включённая исправная цель сохраняет ожидание своей заготовки, даже если
// станок ещё не готов. Нулевой результат только разрешает проверку полезности
// возврата в SELECT_FALLBACK; сам по себе он не требует RETURN_BLANK.
IF SelectMachineForHeldBlank = UINT#0 THEN
	IF (uiCurrentMachine >= FIRST_MACHINE)
	AND (uiCurrentMachine <= LAST_MACHINE) THEN
		IF IsMachineCompatible(
			uiMachine := uiCurrentMachine,
			uiProductType := uiProductType
		) THEN
			SelectMachineForHeldBlank := uiCurrentMachine;
		END_IF;
	END_IF;

	FOR uiMachine := FIRST_MACHINE TO LAST_MACHINE DO
		IF (SelectMachineForHeldBlank = UINT#0)
		AND IsMachineEligible(uiMachine := uiMachine)
		AND (Config.auiMachineType[uiMachine] = uiProductType) THEN
			SelectMachineForHeldBlank := uiMachine;
		END_IF;
	END_FOR;
END_IF;
END_METHOD

METHOD PRIVATE CanReturnHeldBlank : BOOL
VAR
	uiMagazine : UINT; // Магазин следующей операции, независимо от магазина возврата
	uiMachine  : UINT;
	uiType     : UINT;
	uiReservedFreeSlots : UINT; // Возврат занимает один универсальный слот своего магазина
END_VAR
CanReturnHeldBlank := FALSE;

// Для одного типа возврат не открывает нового маршрута. Два груза сначала
// разбираются штатным LOAD/PUT; занятый исправный станок своей заготовки ждём.
IF (Config.uiTypeCount > UINT#1)
AND (Config.uiTypeCount <= UINT#3)
AND stRobotStatus.xBlankAvailable
AND NOT stRobotStatus.xDetailAvailable
AND NOT stRobotStatus.xBusy
AND NOT xStopRequested
AND xMagazineReady
AND (uiBlankPayloadType >= UINT#1)
AND (uiBlankPayloadType <= Config.uiTypeCount) THEN
	IF (stMagazineStatus.stTypeStatus.aiFreeSlot[uiBlankPayloadType] > SINT#0)
	AND (SelectMachineForHeldBlank(
		uiProductType := uiBlankPayloadType,
		uiCurrentMachine := uiSelectedMachine
	) = UINT#0) THEN
		FOR uiMagazine := UINT#1 TO GVL_CELL_SETTINGS.MagazineCount DO
			IF ((uiMagazine = UINT#1) AND xMagazine1Available)
			OR ((uiMagazine = UINT#2) AND xMagazine2Available) THEN
				uiReservedFreeSlots := UINT#0;
				IF uiMagazine = uiActiveMagazine THEN
					uiReservedFreeSlots := UINT#1;
				END_IF;
				FOR uiMachine := FIRST_MACHINE TO LAST_MACHINE DO
					IF IsMachineEligible(uiMachine := uiMachine) THEN
						uiType := Config.auiMachineType[uiMachine];
						IF uiType <> uiBlankPayloadType THEN
							// TAKE освобождает место даже в полной палете. Работающий
							// станок другого типа допускает обычное ожидание его цикла.
							IF (astMagazineStatus[uiMagazine].stTypeStatus.aiBlankSlot[uiType] > SINT#0)
							AND (astMachineStatus[uiMachine].xProcessing
								OR axMachineStartPending[uiMachine]
								OR (astMachineStatus[uiMachine].xCanAcceptService
									AND ((astMachineStatus[uiMachine].ePartState = E_PART_STATE.EMPTY)
										OR astMachineStatus[uiMachine].xServiceRequired))) THEN
								CanReturnHeldBlank := TRUE;
							END_IF;
							// Отдельная выгрузка полезна только для уже готовой детали.
							// Последний свободный слот нельзя занять возвратом и затем
							// выдать UNLOAD без места для этой детали.
							IF astMachineStatus[uiMachine].xCanAcceptService
							AND astMachineStatus[uiMachine].xServiceRequired
							AND (astMachineStatus[uiMachine].ePartState = E_PART_STATE.LOADED)
							AND (astMachineStatus[uiMachine].ePartType = E_PART_TYPE.DETAIL)
							AND (astMagazineStatus[uiMagazine].stTypeStatus.auiFreeCount[uiType] > uiReservedFreeSlots) THEN
								CanReturnHeldBlank := TRUE;
							END_IF;
						END_IF;
					END_IF;
				END_FOR;
			END_IF;
		END_FOR;
	END_IF;
END_IF;
END_METHOD

END_FUNCTION_BLOCK

// Device/Application/FB/F_GEOMETRY_TAKE_DETAIL
FUNCTION F_GEOMETRY_TAKE_DETAIL : BOOL
VAR_INPUT
	uiMachine : UINT;
	uiProductType : UINT;
END_VAR
VAR
	Call : ST_GEOMETRY_CALL;
	EmptyCall : ST_GEOMETRY_CALL;
END_VAR

F_GEOMETRY_TAKE_DETAIL := FALSE;
IF (uiMachine >= UINT#1) AND (uiMachine <= UINT#3) THEN
	// Считаем подтверждённую выгрузку ровно один раз, а не уровень Ready каждый скан.
	// Ожидающая выборка сохраняет счётчик до фактического взятия по FIFO.
	IF (GVL_GEOMETRY_CONTROL.astCalls[uiMachine].uiState <> UINT#1)
	AND GVL_GEOMETRY_CONTROL.xSupported AND GVL_GEOMETRY_CONTROL.xAutoEnabled
	AND (GVL_GEOMETRY_CONTROL.astStatus[1].xEnabled OR GVL_GEOMETRY_CONTROL.astStatus[2].xEnabled) THEN
		GVL_GEOMETRY_CONTROL.auiActiveCount[uiMachine] := MIN(UINT#10000, GVL_GEOMETRY_CONTROL.auiActiveCount[uiMachine] + UINT#1);
		IF GVL_GEOMETRY_CONTROL.auiActiveCount[uiMachine] >= GVL_GEOMETRY_CONTROL.auiPeriod[uiMachine] THEN
			IF (GVL_GEOMETRY_CONTROL.astCalls[uiMachine].uiState <> UINT#2)
			AND (GVL_GEOMETRY_CONTROL.astCalls[uiMachine].uiState <> UINT#3) THEN
				GVL_GEOMETRY_CONTROL.udiNextCallId := GVL_GEOMETRY_CONTROL.udiNextCallId + UDINT#1;
				IF GVL_GEOMETRY_CONTROL.udiNextCallId = UDINT#0 THEN GVL_GEOMETRY_CONTROL.udiNextCallId := UDINT#1; END_IF;
				Call := EmptyCall; Call.udiId := GVL_GEOMETRY_CONTROL.udiNextCallId;
				Call.uiMachine := uiMachine; Call.uiProductType := uiProductType; Call.uiState := UINT#1;
				GVL_GEOMETRY_CONTROL.astCalls[uiMachine] := Call; F_GEOMETRY_EVENT(Call := Call);
			ELSE
				GVL_GEOMETRY_CONTROL.auiActiveCount[uiMachine] := UINT#0;
			END_IF;
		END_IF;
	END_IF;
	// Вызов мог прийти уже после запуска рецепта. Завершаем рецепт, но более
	// поздний вызов оставляем ожидающим следующую деталь, не обгоняя голову FIFO.
	IF (GVL_GEOMETRY_CONTROL.astCalls[uiMachine].uiState = UINT#1)
	AND (F_GEOMETRY_FIRST_CALL() = uiMachine) THEN
		GVL_GEOMETRY_CONTROL.auiActiveCount[uiMachine] := UINT#0;
		GVL_GEOMETRY_CONTROL.astCalls[uiMachine].uiProductType := uiProductType;
		GVL_GEOMETRY_CONTROL.astCalls[uiMachine].uiState := UINT#2;
		F_GEOMETRY_EVENT(Call := GVL_GEOMETRY_CONTROL.astCalls[uiMachine]);
		F_GEOMETRY_TAKE_DETAIL := TRUE;
	END_IF;
END_IF;

END_FUNCTION

// Device/Application/FB/F_GEOMETRY_FIRST_CALL
FUNCTION F_GEOMETRY_FIRST_CALL : UINT
VAR
	uiMachine : UINT;
	udiCallAge : UDINT;
	udiOldestAge : UDINT;
END_VAR

F_GEOMETRY_FIRST_CALL := UINT#0;
udiOldestAge := UDINT#0;
// Только ожидающие вызовы. Готовность станка не меняет его место в FIFO.
FOR uiMachine := UINT#1 TO UINT#3 DO
	IF (GVL_GEOMETRY_CONTROL.astCalls[uiMachine].uiState = UINT#1)
	AND (GVL_GEOMETRY_CONTROL.astCalls[uiMachine].udiId <> UDINT#0) THEN
		// ID монотонный с переходом UDINT_MAX -> 1; нулевой ID пропускается.
		IF GVL_GEOMETRY_CONTROL.udiNextCallId >= GVL_GEOMETRY_CONTROL.astCalls[uiMachine].udiId THEN
			udiCallAge := GVL_GEOMETRY_CONTROL.udiNextCallId - GVL_GEOMETRY_CONTROL.astCalls[uiMachine].udiId;
		ELSE
			udiCallAge := (UDINT#4294967295 - GVL_GEOMETRY_CONTROL.astCalls[uiMachine].udiId)
				+ GVL_GEOMETRY_CONTROL.udiNextCallId;
		END_IF;
		IF (F_GEOMETRY_FIRST_CALL = UINT#0) OR (udiCallAge > udiOldestAge) THEN
			F_GEOMETRY_FIRST_CALL := uiMachine;
			udiOldestAge := udiCallAge;
		END_IF;
	END_IF;
END_FOR;

END_FUNCTION

// Device/Application/FB/FB_FAULT_INJECTOR/FB_CELL_FAULT_INJECTOR
FUNCTION_BLOCK FB_CELL_FAULT_INJECTOR
VAR_INPUT
	Request       : ST_CELL_FAULT_REQUEST; // Запрос локальной ошибки менеджера ячейки
	xOwnerAllowed : BOOL; // Безопасные условия, рассчитанные FB_CELL_MANAGER
END_VAR
VAR_OUTPUT
	xBothGrippers : BOOL; // Одноцикловое противоречивое состояние для штатной проверки
	Status        : ST_FAULT_INJECTION_STATUS; // Состояние источника для HMI
END_VAR
VAR
	rtBothGrippers : R_TRIG; // Фронт команды HMI
END_VAR

rtBothGrippers(CLK := Request.xBothGrippers);
xBothGrippers := FALSE;
Status.xRejected := FALSE;
Status.xAllowed := Request.xEnabled AND xOwnerAllowed;
Status.xBusy := FALSE;
Status.xResetAllowed := FALSE;

IF rtBothGrippers.Q THEN
	IF Status.xAllowed THEN
		xBothGrippers := TRUE;
	ELSE
		Status.xRejected := TRUE;
		Status.udiRejectSequence := Status.udiRejectSequence + UDINT#1;
		IF Status.udiRejectSequence = UDINT#0 THEN
			Status.udiRejectSequence := UDINT#1;
		END_IF;
	END_IF;
END_IF;

Status.xActive := xBothGrippers;

END_FUNCTION_BLOCK

// Device/Application/FB/F_GEOMETRY_SELECT_STATION
FUNCTION F_GEOMETRY_SELECT_STATION : UINT
VAR_INPUT
	xRequireFree : BOOL;
	uiMachine : UINT := UINT#0; // Станок-источник; 0 — общая проверка доступности
END_VAR
VAR
	uiTry : UINT;
	uiStation : UINT;
END_VAR

F_GEOMETRY_SELECT_STATION := UINT#0;
// С1/С2 предпочитают ГК1, С3 — ГК2. История доставок и магазины не участвуют.
uiStation := UINT#1;
IF uiMachine = UINT#3 THEN uiStation := UINT#2; END_IF;
FOR uiTry := UINT#1 TO UINT#2 DO
	// Вторым проверяем другой ГК, если предпочтительный не прошёл допуск.
	IF uiTry = UINT#2 THEN uiStation := UINT#3 - uiStation; END_IF;
	IF (F_GEOMETRY_SELECT_STATION = UINT#0) AND GVL_GEOMETRY_CONTROL.xSupported
	AND GVL_GEOMETRY_CONTROL.astStatus[uiStation].xEnabled
	AND GVL_GEOMETRY_CONTROL.astStatus[uiStation].xConfigured
	AND NOT GVL_GEOMETRY_CONTROL.astStatus[uiStation].xError
	AND (GVL_GEOMETRY_CONTROL.astStatus[uiStation].uiState <> UINT#5) THEN
		IF NOT xRequireFree OR GVL_GEOMETRY_CONTROL.astStatus[uiStation].xReady THEN F_GEOMETRY_SELECT_STATION := uiStation; END_IF;
	END_IF;
END_FOR;

END_FUNCTION

// Device/Application/FB/FB_ALARM_MANAGER
FUNCTION_BLOCK FB_ALARM_MANAGER
VAR_INPUT
	xResetWarnings : BOOL; // Сброс накопленных предупреждений
	astAdditionalCellWarning : ARRAY [1..2] OF ST_WARNING_EVENT; // Конфигуратор и ГК: независимые события источника CELL
END_VAR
VAR_IN_OUT
	Sources : ARRAY [1..19] OF ST_ALARM_SOURCE_DATA; // Старые источники и два ГК
END_VAR
VAR_OUTPUT
	Status : ST_ALARM_STATUS; // Сводный статус журнала
	Events : ARRAY [1..100] OF ST_ALARM_EVENT; // Журнал активных и зафиксированных событий
END_VAR
VAR
	uiWriteIndex : UINT := 1; // Следующая ячейка кольцевого журнала
	udiSequence  : UDINT; // Общий порядковый номер события
	adwPreviousAlarm : ARRAY [1..19] OF DWORD;
	audiPreviousWarning : ARRAY [1..19] OF UDINT;
	audiPreviousAdditionalCellWarning : ARRAY [1..2] OF UDINT;
	uiIndex : UINT; // Индекс источника или события
END_VAR

// Предупреждения подтверждаются только отдельной командой HMI.
// Общий сброс ошибок ячейки не изменяет журнал предупреждений.
IF xResetWarnings THEN
	FOR uiIndex := 1 TO 100 DO
		IF Events[uiIndex].xActive
		AND (Events[uiIndex].eSeverity = E_ALARM_SEVERITY.WARNING) THEN
			Events[uiIndex].xActive := FALSE;
		END_IF;
	END_FOR;
END_IF;

// Менеджер не определяет причины: он регистрирует подготовленные данные владельцев блоков.
FOR uiIndex := 1 TO 19 DO
	UpdateSource(
		eSource := Sources[uiIndex].eSource,
		dwCurrent := Sources[uiIndex].dwAlarmActive,
		xRobotStopRequired := Sources[uiIndex].xRobotStopRequired,
		xGlobalError := Sources[uiIndex].xGlobalError,
		dwPrevious := adwPreviousAlarm[uiIndex]
	);

	IF Sources[uiIndex].stWarning.udiSequence <> audiPreviousWarning[uiIndex] THEN
		IF (Sources[uiIndex].stWarning.udiSequence <> UDINT#0)
		AND (Sources[uiIndex].stWarning.uiCode <> UINT#0) THEN
		AddEvent(
			eSource := Sources[uiIndex].eSource,
			eSeverity := E_ALARM_SEVERITY.WARNING,
			eEffect := E_ALARM_EFFECT.WARNING,
			uiCode := Sources[uiIndex].stWarning.uiCode
		);
		END_IF;
		audiPreviousWarning[uiIndex] := Sources[uiIndex].stWarning.udiSequence;
	END_IF;
END_FOR;

// Общие предупреждения ГК и конфигуратора не изменяют последний код/счётчик
// FB_CELL_MANAGER. Иначе возврат его старого снимка становился новым событием.
// Обрабатываем все каналы в одном вызове: события одного скана не теряются,
// а xResetWarnings не очищает предупреждение, выданное после сброса в этом скане.
FOR uiIndex := UINT#1 TO UINT#2 DO
	IF astAdditionalCellWarning[uiIndex].udiSequence <> audiPreviousAdditionalCellWarning[uiIndex] THEN
		IF (astAdditionalCellWarning[uiIndex].udiSequence <> UDINT#0)
		AND (astAdditionalCellWarning[uiIndex].uiCode <> UINT#0) THEN
			AddEvent(
				eSource := E_ALARM_SOURCE.CELL,
				eSeverity := E_ALARM_SEVERITY.WARNING,
				eEffect := E_ALARM_EFFECT.WARNING,
				uiCode := astAdditionalCellWarning[uiIndex].uiCode
			);
		END_IF;
		audiPreviousAdditionalCellWarning[uiIndex] := astAdditionalCellWarning[uiIndex].udiSequence;
	END_IF;
END_FOR;

Status.uiActiveAlarmCount := 0;
Status.uiActiveWarningCount := 0;
Status.uiHistoryCount := 0;

FOR uiIndex := 1 TO 100 DO
	IF Events[uiIndex].udiSequence <> UDINT#0 THEN
		Status.uiHistoryCount := Status.uiHistoryCount + 1;
	END_IF;
	IF Events[uiIndex].xActive THEN
		IF Events[uiIndex].eSeverity = E_ALARM_SEVERITY.ALARM THEN
			Status.uiActiveAlarmCount := Status.uiActiveAlarmCount + 1;
		ELSE
			Status.uiActiveWarningCount := Status.uiActiveWarningCount + 1;
		END_IF;
	END_IF;
END_FOR;

Status.uiActiveEventCount := Status.uiActiveAlarmCount + Status.uiActiveWarningCount;
Status.xAlarmActive := Status.uiActiveAlarmCount > 0;
Status.xWarningActive := Status.uiActiveWarningCount > 0;

METHOD PRIVATE DeactivateEvent
VAR_INPUT
	eSource : E_ALARM_SOURCE; // Источник аварии
	uiCode  : UINT; // Номер очищенного бита
END_VAR
VAR
	uiIndex : UINT; // Индекс поиска в журнале
END_VAR
FOR uiIndex := 1 TO 100 DO
	IF Events[uiIndex].xActive
	AND (Events[uiIndex].eSeverity = E_ALARM_SEVERITY.ALARM)
	AND (Events[uiIndex].eSource = eSource)
	AND (Events[uiIndex].uiCode = uiCode) THEN
		Events[uiIndex].xActive := FALSE;
	END_IF;
END_FOR;
END_METHOD

METHOD PRIVATE GetAlarmEffect : E_ALARM_EFFECT
VAR_INPUT
	eSource : E_ALARM_SOURCE; // Первичный владелец ошибки
	uiCode : UINT; // Номер бита ошибки владельца
	xRobotStopRequired : BOOL; // Защёлкнутый контекст оборудования требует остановить робота
	xGlobalError : BOOL; // Активна Safety-ошибка ячейки
END_VAR
// Safety имеет абсолютный приоритет над любой частной причиной.
IF xGlobalError THEN
	GetAlarmEffect := E_ALARM_EFFECT.GLOBAL_STOP;

ELSE
CASE eSource OF
	E_ALARM_SOURCE.CELL_SAFETY:
		GetAlarmEffect := E_ALARM_EFFECT.GLOBAL_STOP;

	E_ALARM_SOURCE.CELL:
		CASE uiCode OF
			1: GetAlarmEffect := E_ALARM_EFFECT.ROBOT_STOP; // ERR_ROBOT
			4: GetAlarmEffect := E_ALARM_EFFECT.GLOBAL_STOP; // ERR_GLOBAL_STOP
		ELSE GetAlarmEffect := E_ALARM_EFFECT.EQUIPMENT_STOP;
		END_CASE;

	E_ALARM_SOURCE.MACHINE_1,
	E_ALARM_SOURCE.MACHINE_2,
	E_ALARM_SOURCE.MACHINE_3:
		CASE uiCode OF
			9: GetAlarmEffect := E_ALARM_EFFECT.GLOBAL_STOP; // ERR_SAFETY_STOP
			2, 3, 13, 15, 16, 17, 23: GetAlarmEffect := E_ALARM_EFFECT.ROBOT_STOP;
		ELSE
			IF xRobotStopRequired THEN
				GetAlarmEffect := E_ALARM_EFFECT.ROBOT_STOP;
			ELSE
				GetAlarmEffect := E_ALARM_EFFECT.EQUIPMENT_STOP;
			END_IF;
		END_CASE;

	E_ALARM_SOURCE.MAGAZINE_LOGIC_1,
	E_ALARM_SOURCE.MAGAZINE_LOGIC_2:
		CASE uiCode OF
			5: GetAlarmEffect := E_ALARM_EFFECT.ROBOT_STOP; // ERR_ROBOT
			6: GetAlarmEffect := E_ALARM_EFFECT.GLOBAL_STOP; // ERR_GLOBAL_STOP
		ELSE
			IF xRobotStopRequired THEN
				GetAlarmEffect := E_ALARM_EFFECT.ROBOT_STOP;
			ELSE
				GetAlarmEffect := E_ALARM_EFFECT.EQUIPMENT_STOP;
			END_IF;
		END_CASE;

	E_ALARM_SOURCE.RESERVED_LEGACY_MAGAZINE_AXIS_1,
	E_ALARM_SOURCE.RESERVED_LEGACY_MAGAZINE_AXIS_2,
	E_ALARM_SOURCE.GEOMETRY_1,
	E_ALARM_SOURCE.GEOMETRY_2:
		IF xRobotStopRequired THEN
			GetAlarmEffect := E_ALARM_EFFECT.ROBOT_STOP;
		ELSE
			GetAlarmEffect := E_ALARM_EFFECT.EQUIPMENT_STOP;
		END_IF;

	E_ALARM_SOURCE.ROBOT,
	E_ALARM_SOURCE.AXIS_X,
	E_ALARM_SOURCE.AXIS_Y,
	E_ALARM_SOURCE.AXIS_Z,
	E_ALARM_SOURCE.AXIS_GROUP,
	E_ALARM_SOURCE.MOTION_MANAGER,
	E_ALARM_SOURCE.POINT_MANAGER,
	E_ALARM_SOURCE.GRIPPER:
		GetAlarmEffect := E_ALARM_EFFECT.ROBOT_STOP;

ELSE
	GetAlarmEffect := E_ALARM_EFFECT.EQUIPMENT_STOP;
END_CASE;
END_IF;
END_METHOD

METHOD PRIVATE AddEvent
VAR_INPUT
	eSource   : E_ALARM_SOURCE; // Источник события
	eSeverity : E_ALARM_SEVERITY; // Уровень события
	eEffect   : E_ALARM_EFFECT; // Воздействие события на ячейку
	uiCode    : UINT; // Код события внутри источника
END_VAR
udiSequence := udiSequence + 1;
IF udiSequence = UDINT#0 THEN
	udiSequence := UDINT#1;
END_IF;

Events[uiWriteIndex].udiSequence := udiSequence;
Events[uiWriteIndex].eSeverity := eSeverity;
Events[uiWriteIndex].eEffect := eEffect;
Events[uiWriteIndex].eSource := eSource;
Events[uiWriteIndex].uiCode := uiCode;
Events[uiWriteIndex].xActive := TRUE;

IF uiWriteIndex >= 100 THEN
	uiWriteIndex := 1;
ELSE
	uiWriteIndex := uiWriteIndex + 1;
END_IF;
END_METHOD

METHOD PRIVATE UpdateSource
VAR_INPUT
	eSource   : E_ALARM_SOURCE; // Источник проверяемой маски ошибок
	dwCurrent : DWORD; // Текущая маска ошибок
	xRobotStopRequired : BOOL; // Контекст владельца требует зависимого останова робота
	xGlobalError : BOOL; // Глобальная ошибка активна
END_VAR
VAR_IN_OUT
	dwPrevious : DWORD; // Маска ошибок прошлого цикла
END_VAR
VAR
	dwChanged : DWORD; // Изменившиеся биты
	dwBit     : DWORD; // Маска проверяемого бита
	uiBit     : UINT; // Номер проверяемого бита
END_VAR
dwChanged := dwCurrent XOR dwPrevious;

IF dwChanged <> DWORD#0 THEN
	FOR uiBit := 0 TO 31 DO
		dwBit := SHL(DWORD#1, uiBit);
		IF (dwChanged AND dwBit) <> DWORD#0 THEN
			IF (dwCurrent AND dwBit) <> DWORD#0 THEN
				AddEvent(
					eSource := eSource,
					eSeverity := E_ALARM_SEVERITY.ALARM,
					eEffect := GetAlarmEffect(
						eSource := eSource,
						uiCode := uiBit,
						xRobotStopRequired := xRobotStopRequired,
						xGlobalError := xGlobalError
					),
					uiCode := uiBit
				);
			ELSE
				DeactivateEvent(eSource := eSource, uiCode := uiBit);
			END_IF;
		END_IF;
	END_FOR;
	dwPrevious := dwCurrent;
END_IF;
END_METHOD

END_FUNCTION_BLOCK

// Device/Application/FB/FB_ALARM_HORN
FUNCTION_BLOCK FB_ALARM_HORN
VAR_INPUT
    astSource : ARRAY [1..19] OF ST_ALARM_SOURCE_DATA;
    tDuration : TIME := T#2S;
END_VAR
VAR_OUTPUT
    xSound : BOOL;
END_VAR
VAR
    adwPrevious : ARRAY [1..19] OF DWORD;
    uiSource : UINT;
    xNewAlarm : BOOL;
    xActive : BOOL;
    tLatchedDuration : TIME;
    tonSound : TON;
END_VAR

// Предупреждения не входят в dwAlarmActive. Новая авария другого источника/бита
// тоже запускает звук, даже когда общая xAlarmActive уже была TRUE.
xNewAlarm := FALSE;
FOR uiSource := 1 TO 19 DO
    IF (astSource[uiSource].dwAlarmActive AND NOT adwPrevious[uiSource]) <> DWORD#0 THEN
        xNewAlarm := TRUE;
    END_IF;
    adwPrevious[uiSource] := astSource[uiSource].dwAlarmActive;
END_FOR;
IF tDuration <= T#0MS THEN
    xActive := FALSE;
ELSIF xNewAlarm THEN
    xActive := TRUE;
    tLatchedDuration := tDuration;
    // Сброс и запуск TON в этом же скане: новая авария начинает полный интервал.
    tonSound(IN := FALSE, PT := tLatchedDuration);
END_IF;
tonSound(IN := xActive, PT := tLatchedDuration);
IF tonSound.Q THEN
    xActive := FALSE;
END_IF;
xSound := xActive;

END_FUNCTION_BLOCK

// Device/Application/STATISTIC
PROGRAM STATISTIC
VAR
	fb_Statistic : FB_STATISTIC;
END_VAR

fb_Statistic(
	xStart          := GVL_CELL_MANAGER.Status.xRunning,
	uiSimulationTimeFactor := GVL_CELL_SETTINGS.uiSimulationTimeFactorApplied,
	eActiveAction 	:= GVL_ROBOT.Diag.eActiveAction,
	eActivePoint  	:= GVL_ROBOT.Diag.eActivePoint,
	xBusyMagazine 	:= GVL_MAGAZINE.astStatus[1].xBusy OR GVL_MAGAZINE.astStatus[2].xBusy,
	xBusyMachine_1 	:= GVL_MACHINE.Status[1].xBusy,
	xBusyMachine_2 	:= GVL_MACHINE.Status[2].xBusy,
	xBusyMachine_3 	:= GVL_MACHINE.Status[3].xBusy,
	xCycleActiveMachine_1 	:= GVL_MACHINE.Status[1].stIo.xCycleActive,
	xCycleActiveMachine_2 	:= GVL_MACHINE.Status[2].stIo.xCycleActive,
	xCycleActiveMachine_3 	:= GVL_MACHINE.Status[3].stIo.xCycleActive,
	xBusyRobot 		:=	GVL_ROBOT.Status.xBusy,
	stStatistic     =>  GVL_STATISTIC.stStatistic
);

END_PROGRAM

// Device/Application/FB/FB_STATISTIC/FB_STATISTIC
FUNCTION_BLOCK FB_STATISTIC
VAR_INPUT
	eActiveAction 			: E_ROBOT_ACTION;
	eActivePoint  			: E_POINT_NAME;
	xStart                  : BOOL;
	uiSimulationTimeFactor  : UINT := 1;
	xBusyMagazine       	: BOOL;
	xBusyMachine_1  		: BOOL;
	xBusyMachine_2  		: BOOL;
	xBusyMachine_3  		: BOOL;
	xCycleActiveMachine_1   : BOOL;
	xCycleActiveMachine_2   : BOOL;
	xCycleActiveMachine_3   : BOOL;
	xBusyRobot          	: BOOL;
END_VAR
VAR_OUTPUT
	stStatistic         	: ST_STATISTIC;
END_VAR
VAR
	xInit                   : BOOL;
	xResetStatistics        : BOOL;
	rtSessionStart          : R_TRIG;
	tTotalPLC				: TIME;
	tSessionTime            : TIME;
	tSessionTimeStart       : TIME;
	fbFactorMachine_1 		: FB_CALCULATE;
	fbFactorMachine_2 		: FB_CALCULATE;
	fbFactorMachine_3 		: FB_CALCULATE;
	fbFactorRobot 			: FB_CALCULATE;
	fbAverageMachine_1  	: FB_CALCULATE;
	fbAverageMachine_2  	: FB_CALCULATE;
	fbAverageMachine_3  	: FB_CALCULATE;
	fbAverageMoveMachine_1  : FB_CALCULATE;
	fbAverageMoveMachine_2  : FB_CALCULATE;
	fbAverageMoveMachine_3  : FB_CALCULATE;
	fbAverageMagazine   	: FB_CALCULATE;
END_VAR

rtSessionStart(CLK := xStart);
xResetStatistics := NOT xInit OR rtSessionStart.Q;

IF xResetStatistics THEN
	tSessionTimeStart := TIME();
	xInit := TRUE;
END_IF

tTotalPlc := TIME();
tSessionTime := tTotalPlc - tSessionTimeStart;

fbFactorMachine_1 (
	tTotalPLC := tSessionTime,
	uiSimulationTimeFactor := uiSimulationTimeFactor,
	xMeasure  := xCycleActiveMachine_1,
	xMode := FALSE,
	xReset := xResetStatistics
);

fbFactorMachine_2 (
	tTotalPLC := tSessionTime,
	uiSimulationTimeFactor := uiSimulationTimeFactor,
	xMeasure  := xCycleActiveMachine_2,
	xMode := FALSE,
	xReset := xResetStatistics
);
fbFactorMachine_3 (
	tTotalPLC := tSessionTime,
	uiSimulationTimeFactor := uiSimulationTimeFactor,
	xMeasure  := xCycleActiveMachine_3,
	xMode := FALSE,
	xReset := xResetStatistics
);

fbFactorRobot (
	tTotalPLC := tSessionTime,
	uiSimulationTimeFactor := uiSimulationTimeFactor,
	xMeasure  := xBusyRobot,
	xMode := FALSE,
	xReset := xResetStatistics
);

fbAverageMachine_1(
	uiSimulationTimeFactor := uiSimulationTimeFactor,
	xMeasure  := xBusyMachine_1,
	xMode := TRUE,
	xReset := xResetStatistics
);

fbAverageMachine_2(
	uiSimulationTimeFactor := uiSimulationTimeFactor,
	xMeasure  := xBusyMachine_2,
	xMode := TRUE,
	xReset := xResetStatistics
);

fbAverageMachine_3(
	uiSimulationTimeFactor := uiSimulationTimeFactor,
	xMeasure  := xBusyMachine_3,
	xMode := TRUE,
	xReset := xResetStatistics
);

fbAverageMoveMachine_1(
	uiSimulationTimeFactor := uiSimulationTimeFactor,
	xMeasure  := eActiveAction = E_ROBOT_ACTION.MOVE_TO_POINT AND eActivePoint = E_POINT_NAME.MACHINE_1_ABOVE AND xBusyRobot,
	xMode := TRUE,
	xReset := xResetStatistics
);

fbAverageMoveMachine_2(
	uiSimulationTimeFactor := uiSimulationTimeFactor,
	xMeasure  := eActiveAction = E_ROBOT_ACTION.MOVE_TO_POINT AND eActivePoint = E_POINT_NAME.MACHINE_2_ABOVE AND xBusyRobot,
	xMode := TRUE,
	xReset := xResetStatistics
);

fbAverageMoveMachine_3(
	uiSimulationTimeFactor := uiSimulationTimeFactor,
	xMeasure  := eActiveAction = E_ROBOT_ACTION.MOVE_TO_POINT AND eActivePoint = E_POINT_NAME.MACHINE_3_ABOVE AND xBusyRobot,
	xMode := TRUE,
	xReset := xResetStatistics
);

fbAverageMagazine(
	uiSimulationTimeFactor := uiSimulationTimeFactor,
	xMeasure  := xBusyMagazine,
	xMode := TRUE,
	xReset := xResetStatistics
);


stStatistic.stMachineStat.rLoadCNC_1 := fbFactorMachine_1.rLoadPercent;
stStatistic.stMachineStat.rLoadCNC_2 := fbFactorMachine_2.rLoadPercent;
stStatistic.stMachineStat.rLoadCNC_3 := fbFactorMachine_3.rLoadPercent;
stStatistic.stRobotStat.rRobot       := fbFactorRobot.rLoadPercent;
stStatistic.stRobotStat.tCNC_1       := fbAverageMachine_1.tAverageTime;
stStatistic.stRobotStat.tCNC_2       := fbAverageMachine_2.tAverageTime;
stStatistic.stRobotStat.tCNC_3       := fbAverageMachine_3.tAverageTime;
stStatistic.stRobotStat.tMoveCNC_1   := fbAverageMoveMachine_1.tAverageTime;
stStatistic.stRobotStat.tMoveCNC_2   := fbAverageMoveMachine_2.tAverageTime;
stStatistic.stRobotStat.tMoveCNC_3   := fbAverageMoveMachine_3.tAverageTime;
stStatistic.stRobotStat.tMagazine    := fbAverageMagazine.tAverageTime;

END_FUNCTION_BLOCK

// Device/Application/FB/FB_STATISTIC/FB_CALCULATE
FUNCTION_BLOCK FB_CALCULATE
VAR_INPUT
	xMode          : BOOL;   // Режим работы ФБ (0 - процент загрузки, 1 - среднее время)
	xMeasure 		: BOOL;  // Флаг для измерения загрузки
	tTotalPLC      : TIME;   // Общее время работы ПЛК
	uiSimulationTimeFactor : UINT := 1; // Коэффициент виртуального времени
	xReset         : BOOL;   // Сброс накопленной статистики при старте новой сессии
END_VAR
VAR_OUTPUT
	rLoadPercent 	: REAL;   // Загрузка в процентах
	tAverageTime    : TIME;   // Среднее время
END_VAR
VAR
	uiCount         : UINT;   // Количетво измерений
	rTrig           : R_TRIG; // Фронт сигнала измерения
	fTrig           : F_TRIG; // Спад сигнала измерения
	tStart 			: TIME;   // Время старта замера
	tElapsed        : TIME;   // Измеренное время
	tLastMesured    : TIME;   // Последнее измеренное время
	tTotalBusy      : TIME;   // Общее время загрузки
	tCurrentBusy    : TIME;   // Накопленное время с учётом текущего незавершённого интервала
	tNow            : TIME;   // Текущее системное время
	uiEffectiveTimeFactor : UINT;
	udiScaledTime          : UDINT;
	udiTotalPlcTime        : UDINT;
END_VAR

uiEffectiveTimeFactor := uiSimulationTimeFactor;
IF uiEffectiveTimeFactor < UINT#1 THEN
	uiEffectiveTimeFactor := UINT#1;
ELSIF uiEffectiveTimeFactor > UINT#250 THEN
	uiEffectiveTimeFactor := UINT#250;
END_IF;

tNow := TIME();
rTrig(CLK := xMeasure);
fTrig(CLK := xMeasure);

IF xReset THEN
	uiCount := 0;
	tStart := tNow;
	tElapsed := T#0MS;
	tLastMesured := T#0MS;
	tTotalBusy := T#0MS;
	tCurrentBusy := T#0MS;
	rLoadPercent := 0.0;
	tAverageTime := T#0MS;
ELSE
	IF rTrig.Q THEN
		tStart := tNow;
	END_IF

	IF fTrig.Q THEN
		udiScaledTime := TIME_TO_UDINT(tNow - tStart) * TO_UDINT(uiEffectiveTimeFactor);
		tElapsed := UDINT_TO_TIME(udiScaledTime);
		tTotalBusy := tTotalBusy + tElapsed;
		tLastMesured := tElapsed;
		IF xMode THEN
			uiCount := uiCount + 1;
			tAverageTime := tTotalBusy / uiCount;
		END_IF
	END_IF
END_IF

IF tTotalPLC > T#0S AND NOT xMode THEN
	tCurrentBusy := tTotalBusy;
	IF xMeasure THEN
		udiScaledTime := TIME_TO_UDINT(tNow - tStart) * TO_UDINT(uiEffectiveTimeFactor);
		tCurrentBusy := tCurrentBusy + UDINT_TO_TIME(udiScaledTime);
	END_IF
	udiTotalPlcTime := TIME_TO_UDINT(tTotalPLC) * TO_UDINT(uiEffectiveTimeFactor);
	IF (udiTotalPlcTime > UDINT#0) THEN
		rLoadPercent := UDINT_TO_REAL(TIME_TO_UDINT(tCurrentBusy)) * 100.0
			/ UDINT_TO_REAL(udiTotalPlcTime);
	ELSE
		rLoadPercent := 0.0;
	END_IF;
	IF rLoadPercent > 100.0 THEN
		rLoadPercent := 100.0;
	ELSIF rLoadPercent < 0.0 THEN
		rLoadPercent := 0.0;
	END_IF
ELSIF NOT xMode THEN
	rLoadPercent := 0.0;
END_IF

END_FUNCTION_BLOCK

